(* IEC 61131-3 sources: deprecated-refusr-repo/samples (part 25) *)

(* ---- RND-EXPR_calms-hitch-chips.st ---- *)
(*
This code implements a randomly grown symbolic expression:

((((!(xor(xor(IN37 & (IN27 | ((IN12 & IN24) | (xor(xor(IN9, IN8), IN8)))), (((IN7 & IN10) | (IN4 | IN33)) & IN19) & (xor(xor(!(xor(xor(IN45, IN17), IN10)), !(IN49)), (IN17 & IN40) & (IN49 & IN27)))), (IN29 & (!(xor(xor(IN44, IN27), IN49)))) & IN44))) & (xor(xor((xor(xor(IN25 & ((IN10 | IN28) & IN1), xor(xor(!(!(IN7)), IN13 | (IN39 & IN48)), !(IN32 | IN22))), IN12 & IN3)) & (((!(IN1 & true)) | (IN40 & (!(IN33)))) & ((!(!(IN39))) & ((IN31 | IN24) & IN12))), ((!(IN45)) | ((IN39 | (IN21 | IN31)) | IN2)) | (xor(xor(xor(xor(!(IN20 & IN8), xor(xor(xor(xor(IN3, IN22), IN23), !(IN26)), IN36 & IN23)), !(IN7 | IN30)), (IN12 & (IN40 & IN39)) & (!(IN11 | IN36))), IN48 | IN27))), (!((!(false | IN8)) & ((IN41 & IN46) | (!(IN10))))) & ((!((xor(xor(IN49, IN16), IN2)) | (xor(xor(IN1, IN43), IN14)))) & (!(xor(xor(true & IN26, !(IN43)), xor(xor(IN50, IN38), IN31)))))))) | (((xor(xor(IN15 & (((!(IN16)) & (xor(xor(IN17, IN4), IN20))) & (!(IN23))), (!(xor(xor(false & IN33, xor(xor(IN43, IN26), IN5)), IN34 | IN13))) | (!((xor(xor(IN34, IN42), IN26)) | (!(IN14))))), (((IN10 | IN35) & (IN3 & IN6)) | ((!(IN24)) & (xor(xor(IN26, IN21), IN4)))) | (!(!(IN39 & IN43))))) & (IN6 | ((!(!(xor(xor(IN12, IN16), IN44)))) & IN38))) | (xor(xor(IN25, (xor(xor(xor(xor(!(IN8 & IN48), xor(xor(IN32 | IN43, IN16 | IN16), IN36 | IN46)), xor(xor(IN47, !(IN48)), IN35 | IN43)), xor(xor((IN45 | true) | (!(IN18)), IN13 | (xor(xor(IN5, IN40), IN37))), (!(IN32)) | (!(IN30)))), ((IN6 & IN50) | (IN12 | IN40)) | (xor(xor(!(IN26), xor(xor(IN28, IN10), IN19)), IN30 | IN9)))) & (!(((IN36 & IN40) & (!(IN27))) & (xor(xor(IN36 & true, IN6 | IN2), xor(xor(IN17, IN35), IN35)))))), xor(xor((!(!(IN3 | IN2))) & (!(!(IN13))), IN28), ((!(IN49 & IN49)) | (!(IN7 & IN22))) & (!((IN34 & IN14) & (IN33 | IN12)))))))) & (!(IN3))) & ((!((xor(xor(IN17, !((((IN49 & IN26) | (xor(xor(IN36, IN25), false))) & (xor(xor(IN5 & false, !(IN35)), !(IN50)))) & (!(!(IN6 | IN36))))), !(IN48 & IN8))) & ((xor(xor((!((xor(xor(IN33, IN8), IN42)) | (!(IN38)))) & (xor(xor(!(!(IN31)), xor(xor(IN29, !(IN19)), IN30 & IN32)), xor(xor(IN21, IN19), IN26 | IN33))), (xor(xor((!(IN43)) | (IN50 | IN48), !(!(IN4))), (IN46 | IN17) | (IN30 & IN5))) | ((xor(xor(!(IN13), !(IN13)), xor(xor(IN47, IN28), IN11))) & (xor(xor(!(IN34), IN1 & IN9), IN18 | IN18)))), !(!(!(xor(xor(IN27, IN9), IN50)))))) | (xor(xor(xor(xor(((IN38 | IN16) & (xor(xor(IN41, IN33), IN19))) | (!(xor(xor(IN24, IN1), IN26))), IN22 | ((!(IN32)) | (IN39 & IN2))), ((xor(xor(IN29, IN31), IN5)) & (IN28 | IN27)) & IN20), IN48 & (!((!(IN49)) | (IN30 & IN43)))), IN17 | (((xor(xor(IN21, IN47), IN26)) & (IN28 | false)) | (!(IN31 & false)))))))) & (xor(xor((xor(xor(!((!(!(IN14 & IN46))) & IN35), IN1 | (((!(!(IN20))) & (xor(xor(IN14 & IN29, IN28 & IN20), IN24 & IN18))) & (!(!(IN15 & IN16))))), (xor(xor(((xor(xor(IN14, IN48), IN24)) & (xor(xor(IN5, IN43), IN5))) | ((IN22 | IN46) | (IN44 & IN8)), !((xor(xor(IN50, IN32), IN48)) | (xor(xor(IN28, IN47), IN47)))), (!(xor(xor(IN20, IN39), IN43))) | (!(IN21 & IN17)))) & ((((IN36 | IN24) & (IN9 & IN28)) & IN6) & (true & IN18)))) & ((xor(xor((xor(xor(!(xor(xor(IN44, IN27), IN50)), IN14), IN44)) | (!(!(xor(xor(IN15, IN29), IN24)))), (IN7 & (IN34 | (xor(xor(IN14, IN19), IN41)))) | (((IN10 & IN43) | (IN32 | IN38)) & ((IN5 & IN35) | IN1))), IN43)) | (xor(xor(IN45, xor(xor(true | (!(IN49 | IN18)), IN33 & (!(IN5 & IN13))), IN43)), IN5))), (!((IN23 | ((!(IN45 | IN31)) & IN9)) | (xor(xor(!((IN27 | IN21) & (!(IN26))), !(IN27)), ((IN48 & IN48) & (xor(xor(IN37, IN41), IN13))) & IN49)))) | (((!(((!(IN15)) | (xor(xor(IN1, IN25), IN6))) | IN46)) | IN13) & ((IN18 | (xor(xor(IN14 & (!(IN35)), xor(xor(xor(xor(IN40, IN41), IN23), xor(xor(IN6, IN18), IN22)), IN10)), IN35))) | (!(((IN34 & IN11) & (IN46 & IN43)) & (xor(xor(IN31, IN25 | IN32), xor(xor(IN35, IN11), IN9)))))))), !(((xor(xor(xor(xor(IN39, IN42 | (xor(xor(IN33, IN4), IN29))), IN24 & (!(IN45))), (xor(xor(!(IN11), IN39 & false), IN35)) & ((xor(xor(IN12, IN35), IN44)) & IN30)), xor(xor(IN23, !(!(IN25))), !(IN25 & IN14)))) & (IN24 | ((xor(xor(IN4, !(IN27)), IN28 | IN44)) | (xor(xor(IN44 & IN22, IN44 | IN50), IN44))))) | (!((xor(xor(!(IN23), (xor(xor(IN24, IN35), IN27)) & (IN27 | IN14)), (!(IN37)) & (!(IN27)))) & ((xor(xor(IN24 & IN33, IN3), !(IN16))) & ((IN12 | IN39) & IN25))))))))

*)

FUNCTION_BLOCK F_CollectInput
  VAR_IN_OUT
      Data : ARRAY[1..50] OF BOOL;
  END_VAR
  VAR_INPUT
      TICK  : BOOL := 0;
      IN1   : BOOL := 0;
      IN2   : BOOL := 0;
      IN3   : BOOL := 0;
      IN4   : BOOL := 0;
      IN5   : BOOL := 0;
      RESET : BOOL := FALSE;
  END_VAR
  VAR_OUTPUT
      Finished : BOOL;
  END_VAR
  VAR
      j    : USINT := 1;
      tock : BOOL  := 0;
  END_VAR
  IF NOT RESET AND tock = NOT TICK THEN
      Data[j]   := IN1;
      Data[j+1] := IN2;
      Data[j+2] := IN3;
      Data[j+3] := IN4;
      Data[j+4] := IN5;
      j := j + 5;
      tock := TICK;
  ELSE
      j := 1;
      tock := 0;
  END_IF;
  Finished := (j > 50);
END_FUNCTION_BLOCK

PROGRAM Boiler
  VAR
    Data  : ARRAY[1..50] OF BOOL;
    Ready : BOOL;
    CollectInput : F_CollectInput;
  END_VAR
  VAR
    TICK     AT %IX1.0 : BOOL;
    IN1      AT %IX0.3 : BOOL;
    IN2      AT %IX0.4 : BOOL;
    IN3      AT %IX0.5 : BOOL;
    IN4      AT %IX0.6 : BOOL;
    IN5      AT %IX0.7 : BOOL;
    OutReady AT %QX0.0 : BOOL := FALSE;
    FeedNext AT %QX0.1 : BOOL := FALSE;
    Out      AT %QX0.2 : BOOL;
  END_VAR
  CollectInput(TICK:=TICK, IN1:=IN1, IN2:=IN2, IN3:=IN3, IN4:=IN4, IN5:=IN5);
  Ready := CollectInput.Finished;
  FeedNext := 1;
  IF Ready THEN
    Out := (((((NOT (((Data[37] AND (Data[27] OR ((Data[12] AND Data[24]) OR ((Data[9] XOR Data[8]) XOR Data[8])))) XOR ((((Data[7] AND Data[10]) OR (Data[4] OR Data[33])) AND Data[19]) AND (((NOT ((Data[45] XOR Data[17]) XOR Data[10])) XOR (NOT Data[49])) XOR ((Data[17] AND Data[40]) AND (Data[49] AND Data[27]))))) XOR ((Data[29] AND (NOT ((Data[44] XOR Data[27]) XOR Data[49]))) AND Data[44]))) AND ((((((Data[25] AND ((Data[10] OR Data[28]) AND Data[1])) XOR (((NOT (NOT Data[7])) XOR (Data[13] OR (Data[39] AND Data[48]))) XOR (NOT (Data[32] OR Data[22])))) XOR (Data[12] AND Data[3])) AND (((NOT (Data[1] AND TRUE)) OR (Data[40] AND (NOT Data[33]))) AND ((NOT (NOT Data[39])) AND ((Data[31] OR Data[24]) AND Data[12])))) XOR (((NOT Data[45]) OR ((Data[39] OR (Data[21] OR Data[31])) OR Data[2])) OR (((((NOT (Data[20] AND Data[8])) XOR ((((Data[3] XOR Data[22]) XOR Data[23]) XOR (NOT Data[26])) XOR (Data[36] AND Data[23]))) XOR (NOT (Data[7] OR Data[30]))) XOR ((Data[12] AND (Data[40] AND Data[39])) AND (NOT (Data[11] OR Data[36])))) XOR (Data[48] OR Data[27])))) XOR ((NOT ((NOT (FALSE OR Data[8])) AND ((Data[41] AND Data[46]) OR (NOT Data[10])))) AND ((NOT (((Data[49] XOR Data[16]) XOR Data[2]) OR ((Data[1] XOR Data[43]) XOR Data[14]))) AND (NOT (((TRUE AND Data[26]) XOR (NOT Data[43])) XOR ((Data[50] XOR Data[38]) XOR Data[31]))))))) OR (((((Data[15] AND (((NOT Data[16]) AND ((Data[17] XOR Data[4]) XOR Data[20])) AND (NOT Data[23]))) XOR ((NOT (((FALSE AND Data[33]) XOR ((Data[43] XOR Data[26]) XOR Data[5])) XOR (Data[34] OR Data[13]))) OR (NOT (((Data[34] XOR Data[42]) XOR Data[26]) OR (NOT Data[14]))))) XOR ((((Data[10] OR Data[35]) AND (Data[3] AND Data[6])) OR ((NOT Data[24]) AND ((Data[26] XOR Data[21]) XOR Data[4]))) OR (NOT (NOT (Data[39] AND Data[43]))))) AND (Data[6] OR ((NOT (NOT ((Data[12] XOR Data[16]) XOR Data[44]))) AND Data[38]))) OR ((Data[25] XOR ((((((NOT (Data[8] AND Data[48])) XOR (((Data[32] OR Data[43]) XOR (Data[16] OR Data[16])) XOR (Data[36] OR Data[46]))) XOR ((Data[47] XOR (NOT Data[48])) XOR (Data[35] OR Data[43]))) XOR ((((Data[45] OR TRUE) OR (NOT Data[18])) XOR (Data[13] OR ((Data[5] XOR Data[40]) XOR Data[37]))) XOR ((NOT Data[32]) OR (NOT Data[30])))) XOR (((Data[6] AND Data[50]) OR (Data[12] OR Data[40])) OR (((NOT Data[26]) XOR ((Data[28] XOR Data[10]) XOR Data[19])) XOR (Data[30] OR Data[9])))) AND (NOT (((Data[36] AND Data[40]) AND (NOT Data[27])) AND (((Data[36] AND TRUE) XOR (Data[6] OR Data[2])) XOR ((Data[17] XOR Data[35]) XOR Data[35])))))) XOR ((((NOT (NOT (Data[3] OR Data[2]))) AND (NOT (NOT Data[13]))) XOR Data[28]) XOR (((NOT (Data[49] AND Data[49])) OR (NOT (Data[7] AND Data[22]))) AND (NOT ((Data[34] AND Data[14]) AND (Data[33] OR Data[12])))))))) AND (NOT Data[3])) AND ((NOT (((Data[17] XOR (NOT ((((Data[49] AND Data[26]) OR ((Data[36] XOR Data[25]) XOR FALSE)) AND (((Data[5] AND FALSE) XOR (NOT Data[35])) XOR (NOT Data[50]))) AND (NOT (NOT (Data[6] OR Data[36])))))) XOR (NOT (Data[48] AND Data[8]))) AND (((((NOT (((Data[33] XOR Data[8]) XOR Data[42]) OR (NOT Data[38]))) AND (((NOT (NOT Data[31])) XOR ((Data[29] XOR (NOT Data[19])) XOR (Data[30] AND Data[32]))) XOR ((Data[21] XOR Data[19]) XOR (Data[26] OR Data[33])))) XOR (((((NOT Data[43]) OR (Data[50] OR Data[48])) XOR (NOT (NOT Data[4]))) XOR ((Data[46] OR Data[17]) OR (Data[30] AND Data[5]))) OR ((((NOT Data[13]) XOR (NOT Data[13])) XOR ((Data[47] XOR Data[28]) XOR Data[11])) AND (((NOT Data[34]) XOR (Data[1] AND Data[9])) XOR (Data[18] OR Data[18]))))) XOR (NOT (NOT (NOT ((Data[27] XOR Data[9]) XOR Data[50]))))) OR (((((((Data[38] OR Data[16]) AND ((Data[41] XOR Data[33]) XOR Data[19])) OR (NOT ((Data[24] XOR Data[1]) XOR Data[26]))) XOR (Data[22] OR ((NOT Data[32]) OR (Data[39] AND Data[2])))) XOR ((((Data[29] XOR Data[31]) XOR Data[5]) AND (Data[28] OR Data[27])) AND Data[20])) XOR (Data[48] AND (NOT ((NOT Data[49]) OR (Data[30] AND Data[43]))))) XOR (Data[17] OR ((((Data[21] XOR Data[47]) XOR Data[26]) AND (Data[28] OR FALSE)) OR (NOT (Data[31] AND FALSE)))))))) AND ((((((NOT ((NOT (NOT (Data[14] AND Data[46]))) AND Data[35])) XOR (Data[1] OR (((NOT (NOT Data[20])) AND (((Data[14] AND Data[29]) XOR (Data[28] AND Data[20])) XOR (Data[24] AND Data[18]))) AND (NOT (NOT (Data[15] AND Data[16])))))) XOR (((((((Data[14] XOR Data[48]) XOR Data[24]) AND ((Data[5] XOR Data[43]) XOR Data[5])) OR ((Data[22] OR Data[46]) OR (Data[44] AND Data[8]))) XOR (NOT (((Data[50] XOR Data[32]) XOR Data[48]) OR ((Data[28] XOR Data[47]) XOR Data[47])))) XOR ((NOT ((Data[20] XOR Data[39]) XOR Data[43])) OR (NOT (Data[21] AND Data[17])))) AND ((((Data[36] OR Data[24]) AND (Data[9] AND Data[28])) AND Data[6]) AND (TRUE AND Data[18])))) AND (((((((NOT ((Data[44] XOR Data[27]) XOR Data[50])) XOR Data[14]) XOR Data[44]) OR (NOT (NOT ((Data[15] XOR Data[29]) XOR Data[24])))) XOR ((Data[7] AND (Data[34] OR ((Data[14] XOR Data[19]) XOR Data[41]))) OR (((Data[10] AND Data[43]) OR (Data[32] OR Data[38])) AND ((Data[5] AND Data[35]) OR Data[1])))) XOR Data[43]) OR ((Data[45] XOR (((TRUE OR (NOT (Data[49] OR Data[18]))) XOR (Data[33] AND (NOT (Data[5] AND Data[13])))) XOR Data[43])) XOR Data[5]))) XOR ((NOT ((Data[23] OR ((NOT (Data[45] OR Data[31])) AND Data[9])) OR (((NOT ((Data[27] OR Data[21]) AND (NOT Data[26]))) XOR (NOT Data[27])) XOR (((Data[48] AND Data[48]) AND ((Data[37] XOR Data[41]) XOR Data[13])) AND Data[49])))) OR (((NOT (((NOT Data[15]) OR ((Data[1] XOR Data[25]) XOR Data[6])) OR Data[46])) OR Data[13]) AND ((Data[18] OR (((Data[14] AND (NOT Data[35])) XOR ((((Data[40] XOR Data[41]) XOR Data[23]) XOR ((Data[6] XOR Data[18]) XOR Data[22])) XOR Data[10])) XOR Data[35])) OR (NOT (((Data[34] AND Data[11]) AND (Data[46] AND Data[43])) AND ((Data[31] XOR (Data[25] OR Data[32])) XOR ((Data[35] XOR Data[11]) XOR Data[9])))))))) XOR (NOT ((((((Data[39] XOR (Data[42] OR ((Data[33] XOR Data[4]) XOR Data[29]))) XOR (Data[24] AND (NOT Data[45]))) XOR ((((NOT Data[11]) XOR (Data[39] AND FALSE)) XOR Data[35]) AND (((Data[12] XOR Data[35]) XOR Data[44]) AND Data[30]))) XOR ((Data[23] XOR (NOT (NOT Data[25]))) XOR (NOT (Data[25] AND Data[14])))) AND (Data[24] OR (((Data[4] XOR (NOT Data[27])) XOR (Data[28] OR Data[44])) OR (((Data[44] AND Data[22]) XOR (Data[44] OR Data[50])) XOR Data[44])))) OR (NOT ((((NOT Data[23]) XOR (((Data[24] XOR Data[35]) XOR Data[27]) AND (Data[27] OR Data[14]))) XOR ((NOT Data[37]) AND (NOT Data[27]))) AND ((((Data[24] AND Data[33]) XOR Data[3]) XOR (NOT Data[16])) AND ((Data[12] OR Data[39]) AND Data[25])))))))));
    OutReady := 1;
    CollectInput(RESET:=TRUE);
  END_IF;
END_PROGRAM

CONFIGURATION Config0
  RESOURCE Res0 ON PLC
    TASK task0(INTERVAL := T#20ms,PRIORITY := 0);
    PROGRAM instance0 WITH task0 : Boiler;
  END_RESOURCE
END_CONFIGURATION

(* ---- RND-EXPR_celeb-candy-degas.st ---- *)
(*
This code implements a randomly grown symbolic expression:

!(xor(xor(!(!(((IN43 & ((xor(xor(IN28 | IN19, !(IN27)), IN33 | IN34)) & (xor(xor(xor(xor(IN27, IN17), IN17), xor(xor(true, IN6), IN43)), xor(xor(IN12, IN24), IN27))))) | IN22) & ((!(xor(xor(IN48, true), IN11))) | (((!(IN32)) | (!(IN3 | IN3))) | ((!(IN10)) | ((IN29 | IN6) | IN19)))))), xor(xor(xor(xor(IN26, !(IN24)), ((IN50 | ((xor(xor(IN4 & IN32, xor(xor(IN29, IN44), IN1)), IN25 & IN41)) | ((IN17 | IN36) & (xor(xor(IN10, IN2), IN16))))) & ((!(!(IN10))) | (!((!(IN48)) | (IN8 | IN19))))) | (!(!(((IN1 | IN6) | IN48) | (IN15 & IN7))))), ((xor(xor(xor(xor((xor(xor(!(IN39), !(IN1)), IN33 | IN10)) | IN5, xor(xor((IN21 | IN15) & (xor(xor(IN35, IN25), IN41)), (IN18 | IN2) & IN21), (IN2 | IN3) & (!(IN39)))), xor(xor((IN36 | IN33) | (!(IN14)), !(!(IN39))), !(IN16 & IN8))), IN15), (xor(xor(xor(xor(IN6 | IN24, xor(xor(IN49, IN14), IN21)), xor(xor(IN13, IN16), IN43)), !(xor(xor(IN23, IN10), IN19))), xor(xor(IN6 | IN31, xor(xor(IN40, IN38), IN29)), IN43))) & ((IN38 | (!(IN28))) | ((xor(xor(IN33, IN34), IN36)) & IN13)))) | IN42) | (((xor(xor((xor(xor(IN4, xor(xor(IN6, IN6), IN31)), !(IN21))) | (!(xor(xor(IN21, false), IN15))), IN17), ((xor(xor(false, IN5), IN47)) & (xor(xor(IN49, IN19), IN41))) & (xor(xor(!(IN38), IN8 | IN34), IN15 & IN16)))) | IN18) & ((IN38 & (IN28 & IN1)) | (xor(xor((IN10 | (!(IN33))) | IN45, (!(IN6 & IN5)) & ((!(IN3)) | IN19)), xor(xor(xor(xor(!(IN28), IN16 | IN32), IN2 | IN9), (IN39 | IN36) & (!(IN41))), (!(IN26)) | (!(IN47)))))))), xor(xor(!(((((IN14 | false) & IN34) & (IN23 & (IN13 | IN3))) & (((IN45 & IN1) | (xor(xor(IN22, IN35), IN4))) | (IN2 & IN25))) | IN26), xor(xor(xor(xor((IN2 & (xor(xor(xor(xor(IN4, IN28), IN34), IN3 & IN28), IN24 | IN22))) | IN16, (xor(xor(!(IN26 & IN50), !(IN13 | IN37)), !(IN35))) | (((!(IN35)) & IN24) & (!(IN24 & IN12)))), xor(xor(!((!(IN10)) | (IN9 | IN28)), ((IN35 | IN46) & IN4) | (xor(xor(false, xor(xor(IN22, IN24), IN1)), IN22 | IN21))), ((IN29 & IN33) | (xor(xor(false, IN45), IN26))) | IN30)), !(IN19)), xor(xor(false, !((xor(xor(IN22 | IN45, xor(xor(IN12, true), IN19)), IN35 & IN24)) | (!(IN46)))), IN50))), IN39))), xor(xor(IN12 & (xor(xor(!(xor(xor(((xor(xor(IN31, IN35), IN20)) & (!(IN37))) & ((xor(xor(IN15, IN38), IN12)) & (xor(xor(IN19, IN42), IN31))), ((IN9 & IN29) | (!(IN16))) & IN5), ((xor(xor(IN21, IN25), IN21)) | (IN21 | IN17)) & (!(!(IN42))))), xor(xor((xor(xor(IN12, !(xor(xor(IN48, true), IN39))), (IN21 | IN43) | (IN12 | true))) | ((xor(xor(IN31 | IN44, IN18 & IN48), xor(xor(IN11, IN35), IN21))) & (xor(xor(xor(xor(IN25, IN40), IN10), IN13 & true), xor(xor(IN47, IN22), IN21)))), (xor(xor((!(IN36)) & (IN29 & IN15), IN35), IN46)) & (!(IN32))), !(!((!(IN27)) & (!(IN36)))))), (!(((IN1 & IN21) | (!(IN45))) | ((IN23 & IN32) | IN41))) & (xor(xor(xor(xor(IN40, (!(IN32)) & (IN20 | IN20)), xor(xor(xor(xor(IN26, IN20), IN50), IN8 & IN49), IN4 & IN21)), ((xor(xor(IN25, IN6), IN39)) & (IN10 & IN16)) & (xor(xor(IN14 & IN33, IN3 & IN21), IN28 | IN18))), IN13)))), xor(xor(xor(xor(!((!(xor(xor(IN29 & IN49, IN32), xor(xor(IN15, IN21), IN3)))) | (!(IN49 & (xor(xor(IN23, IN40), IN49))))), (xor(xor(((!(IN49)) & (IN28 & IN26)) & IN23, ((IN43 & IN42) | IN39) & (!(IN38 | IN22))), (!(IN17)) & IN50)) & ((xor(xor(xor(xor(xor(xor(IN50, IN5), IN38), xor(xor(IN49, IN32), IN31)), !(IN18)), IN11), (!(IN6)) | IN38)) & IN48)), IN50 & IN22), ((xor(xor(IN31 & true, (!(IN47 & IN18)) | (!(!(IN48)))), (!(!(IN50))) | IN28)) | ((!((IN7 | IN24) | (IN4 | IN44))) | (xor(xor(!(IN9), IN39), (false & IN12) | (IN26 & IN50))))) & IN35), !((!(xor(xor(IN7, (!(IN38)) & (IN38 | IN17)), xor(xor(xor(xor(IN49, IN21), IN35), IN17 & IN21), xor(xor(IN45, IN26), IN29))))) | ((IN36 & (xor(xor(xor(xor(IN11, IN31), IN32), IN46 & IN49), !(IN2)))) & (!(!(IN24))))))), xor(xor(xor(xor(!(IN1 & IN12), (!(xor(xor(xor(xor(!(IN44), IN35), IN41 | IN16), xor(xor(IN39 & IN2, !(IN19)), IN25)), !(IN21)))) | ((((xor(xor(IN27, IN33), false)) & IN29) | ((IN4 & IN18) | (IN2 | IN36))) & IN46)), (IN23 | (!(IN13))) & (!((true & (IN42 & IN20)) | (xor(xor(!(IN12), IN7 | true), IN1 | IN14))))), IN21), !(!(IN29))))))

*)

FUNCTION_BLOCK F_CollectInput
  VAR_IN_OUT
      Data : ARRAY[1..50] OF BOOL;
  END_VAR
  VAR_INPUT
      TICK  : BOOL := 0;
      IN1   : BOOL := 0;
      IN2   : BOOL := 0;
      IN3   : BOOL := 0;
      IN4   : BOOL := 0;
      IN5   : BOOL := 0;
      RESET : BOOL := FALSE;
  END_VAR
  VAR_OUTPUT
      Finished : BOOL;
  END_VAR
  VAR
      j    : USINT := 1;
      tock : BOOL  := 0;
  END_VAR
  IF NOT RESET AND tock = NOT TICK THEN
      Data[j]   := IN1;
      Data[j+1] := IN2;
      Data[j+2] := IN3;
      Data[j+3] := IN4;
      Data[j+4] := IN5;
      j := j + 5;
      tock := TICK;
  ELSE
      j := 1;
      tock := 0;
  END_IF;
  Finished := (j > 50);
END_FUNCTION_BLOCK

PROGRAM Boiler
  VAR
    Data  : ARRAY[1..50] OF BOOL;
    Ready : BOOL;
    CollectInput : F_CollectInput;
  END_VAR
  VAR
    TICK     AT %IX1.0 : BOOL;
    IN1      AT %IX0.3 : BOOL;
    IN2      AT %IX0.4 : BOOL;
    IN3      AT %IX0.5 : BOOL;
    IN4      AT %IX0.6 : BOOL;
    IN5      AT %IX0.7 : BOOL;
    OutReady AT %QX0.0 : BOOL := FALSE;
    FeedNext AT %QX0.1 : BOOL := FALSE;
    Out      AT %QX0.2 : BOOL;
  END_VAR
  CollectInput(TICK:=TICK, IN1:=IN1, IN2:=IN2, IN3:=IN3, IN4:=IN4, IN5:=IN5);
  Ready := CollectInput.Finished;
  FeedNext := 1;
  IF Ready THEN
    Out := (NOT (((NOT (NOT (((Data[43] AND ((((Data[28] OR Data[19]) XOR (NOT Data[27])) XOR (Data[33] OR Data[34])) AND ((((Data[27] XOR Data[17]) XOR Data[17]) XOR ((TRUE XOR Data[6]) XOR Data[43])) XOR ((Data[12] XOR Data[24]) XOR Data[27])))) OR Data[22]) AND ((NOT ((Data[48] XOR TRUE) XOR Data[11])) OR (((NOT Data[32]) OR (NOT (Data[3] OR Data[3]))) OR ((NOT Data[10]) OR ((Data[29] OR Data[6]) OR Data[19]))))))) XOR ((((Data[26] XOR (NOT Data[24])) XOR (((Data[50] OR ((((Data[4] AND Data[32]) XOR ((Data[29] XOR Data[44]) XOR Data[1])) XOR (Data[25] AND Data[41])) OR ((Data[17] OR Data[36]) AND ((Data[10] XOR Data[2]) XOR Data[16])))) AND ((NOT (NOT Data[10])) OR (NOT ((NOT Data[48]) OR (Data[8] OR Data[19]))))) OR (NOT (NOT (((Data[1] OR Data[6]) OR Data[48]) OR (Data[15] AND Data[7])))))) XOR ((((((((((NOT Data[39]) XOR (NOT Data[1])) XOR (Data[33] OR Data[10])) OR Data[5]) XOR ((((Data[21] OR Data[15]) AND ((Data[35] XOR Data[25]) XOR Data[41])) XOR ((Data[18] OR Data[2]) AND Data[21])) XOR ((Data[2] OR Data[3]) AND (NOT Data[39])))) XOR ((((Data[36] OR Data[33]) OR (NOT Data[14])) XOR (NOT (NOT Data[39]))) XOR (NOT (Data[16] AND Data[8])))) XOR Data[15]) XOR ((((((Data[6] OR Data[24]) XOR ((Data[49] XOR Data[14]) XOR Data[21])) XOR ((Data[13] XOR Data[16]) XOR Data[43])) XOR (NOT ((Data[23] XOR Data[10]) XOR Data[19]))) XOR (((Data[6] OR Data[31]) XOR ((Data[40] XOR Data[38]) XOR Data[29])) XOR Data[43])) AND ((Data[38] OR (NOT Data[28])) OR (((Data[33] XOR Data[34]) XOR Data[36]) AND Data[13])))) OR Data[42]) OR (((((((Data[4] XOR ((Data[6] XOR Data[6]) XOR Data[31])) XOR (NOT Data[21])) OR (NOT ((Data[21] XOR FALSE) XOR Data[15]))) XOR Data[17]) XOR ((((FALSE XOR Data[5]) XOR Data[47]) AND ((Data[49] XOR Data[19]) XOR Data[41])) AND (((NOT Data[38]) XOR (Data[8] OR Data[34])) XOR (Data[15] AND Data[16])))) OR Data[18]) AND ((Data[38] AND (Data[28] AND Data[1])) OR ((((Data[10] OR (NOT Data[33])) OR Data[45]) XOR ((NOT (Data[6] AND Data[5])) AND ((NOT Data[3]) OR Data[19]))) XOR (((((NOT Data[28]) XOR (Data[16] OR Data[32])) XOR (Data[2] OR Data[9])) XOR ((Data[39] OR Data[36]) AND (NOT Data[41]))) XOR ((NOT Data[26]) OR (NOT Data[47])))))))) XOR (((NOT (((((Data[14] OR FALSE) AND Data[34]) AND (Data[23] AND (Data[13] OR Data[3]))) AND (((Data[45] AND Data[1]) OR ((Data[22] XOR Data[35]) XOR Data[4])) OR (Data[2] AND Data[25]))) OR Data[26])) XOR ((((((Data[2] AND ((((Data[4] XOR Data[28]) XOR Data[34]) XOR (Data[3] AND Data[28])) XOR (Data[24] OR Data[22]))) OR Data[16]) XOR ((((NOT (Data[26] AND Data[50])) XOR (NOT (Data[13] OR Data[37]))) XOR (NOT Data[35])) OR (((NOT Data[35]) AND Data[24]) AND (NOT (Data[24] AND Data[12]))))) XOR (((NOT ((NOT Data[10]) OR (Data[9] OR Data[28]))) XOR (((Data[35] OR Data[46]) AND Data[4]) OR ((FALSE XOR ((Data[22] XOR Data[24]) XOR Data[1])) XOR (Data[22] OR Data[21])))) XOR (((Data[29] AND Data[33]) OR ((FALSE XOR Data[45]) XOR Data[26])) OR Data[30]))) XOR (NOT Data[19])) XOR ((FALSE XOR (NOT ((((Data[22] OR Data[45]) XOR ((Data[12] XOR TRUE) XOR Data[19])) XOR (Data[35] AND Data[24])) OR (NOT Data[46])))) XOR Data[50]))) XOR Data[39]))) XOR (((Data[12] AND (((NOT ((((((Data[31] XOR Data[35]) XOR Data[20]) AND (NOT Data[37])) AND (((Data[15] XOR Data[38]) XOR Data[12]) AND ((Data[19] XOR Data[42]) XOR Data[31]))) XOR (((Data[9] AND Data[29]) OR (NOT Data[16])) AND Data[5])) XOR ((((Data[21] XOR Data[25]) XOR Data[21]) OR (Data[21] OR Data[17])) AND (NOT (NOT Data[42]))))) XOR (((((Data[12] XOR (NOT ((Data[48] XOR TRUE) XOR Data[39]))) XOR ((Data[21] OR Data[43]) OR (Data[12] OR TRUE))) OR ((((Data[31] OR Data[44]) XOR (Data[18] AND Data[48])) XOR ((Data[11] XOR Data[35]) XOR Data[21])) AND ((((Data[25] XOR Data[40]) XOR Data[10]) XOR (Data[13] AND TRUE)) XOR ((Data[47] XOR Data[22]) XOR Data[21])))) XOR (((((NOT Data[36]) AND (Data[29] AND Data[15])) XOR Data[35]) XOR Data[46]) AND (NOT Data[32]))) XOR (NOT (NOT ((NOT Data[27]) AND (NOT Data[36])))))) XOR ((NOT (((Data[1] AND Data[21]) OR (NOT Data[45])) OR ((Data[23] AND Data[32]) OR Data[41]))) AND ((((Data[40] XOR ((NOT Data[32]) AND (Data[20] OR Data[20]))) XOR ((((Data[26] XOR Data[20]) XOR Data[50]) XOR (Data[8] AND Data[49])) XOR (Data[4] AND Data[21]))) XOR ((((Data[25] XOR Data[6]) XOR Data[39]) AND (Data[10] AND Data[16])) AND (((Data[14] AND Data[33]) XOR (Data[3] AND Data[21])) XOR (Data[28] OR Data[18])))) XOR Data[13])))) XOR (((((NOT ((NOT (((Data[29] AND Data[49]) XOR Data[32]) XOR ((Data[15] XOR Data[21]) XOR Data[3]))) OR (NOT (Data[49] AND ((Data[23] XOR Data[40]) XOR Data[49]))))) XOR ((((((NOT Data[49]) AND (Data[28] AND Data[26])) AND Data[23]) XOR (((Data[43] AND Data[42]) OR Data[39]) AND (NOT (Data[38] OR Data[22])))) XOR ((NOT Data[17]) AND Data[50])) AND (((((((Data[50] XOR Data[5]) XOR Data[38]) XOR ((Data[49] XOR Data[32]) XOR Data[31])) XOR (NOT Data[18])) XOR Data[11]) XOR ((NOT Data[6]) OR Data[38])) AND Data[48]))) XOR (Data[50] AND Data[22])) XOR (((((Data[31] AND TRUE) XOR ((NOT (Data[47] AND Data[18])) OR (NOT (NOT Data[48])))) XOR ((NOT (NOT Data[50])) OR Data[28])) OR ((NOT ((Data[7] OR Data[24]) OR (Data[4] OR Data[44]))) OR (((NOT Data[9]) XOR Data[39]) XOR ((FALSE AND Data[12]) OR (Data[26] AND Data[50]))))) AND Data[35])) XOR (NOT ((NOT ((Data[7] XOR ((NOT Data[38]) AND (Data[38] OR Data[17]))) XOR ((((Data[49] XOR Data[21]) XOR Data[35]) XOR (Data[17] AND Data[21])) XOR ((Data[45] XOR Data[26]) XOR Data[29])))) OR ((Data[36] AND ((((Data[11] XOR Data[31]) XOR Data[32]) XOR (Data[46] AND Data[49])) XOR (NOT Data[2]))) AND (NOT (NOT Data[24]))))))) XOR (((((NOT (Data[1] AND Data[12])) XOR ((NOT (((((NOT Data[44]) XOR Data[35]) XOR (Data[41] OR Data[16])) XOR (((Data[39] AND Data[2]) XOR (NOT Data[19])) XOR Data[25])) XOR (NOT Data[21]))) OR (((((Data[27] XOR Data[33]) XOR FALSE) AND Data[29]) OR ((Data[4] AND Data[18]) OR (Data[2] OR Data[36]))) AND Data[46]))) XOR ((Data[23] OR (NOT Data[13])) AND (NOT ((TRUE AND (Data[42] AND Data[20])) OR (((NOT Data[12]) XOR (Data[7] OR TRUE)) XOR (Data[1] OR Data[14])))))) XOR Data[21]) XOR (NOT (NOT Data[29]))))));
    OutReady := 1;
    CollectInput(RESET:=TRUE);
  END_IF;
END_PROGRAM

CONFIGURATION Config0
  RESOURCE Res0 ON PLC
    TASK task0(INTERVAL := T#20ms,PRIORITY := 0);
    PROGRAM instance0 WITH task0 : Boiler;
  END_RESOURCE
END_CONFIGURATION

(* ---- RND-EXPR_endue-lawns-artsy.st ---- *)
(*
This code implements a randomly grown symbolic expression:

xor(xor(xor(xor(!(xor(xor(IN45, xor(xor((((xor(xor(IN19 & IN49, IN3 & IN10), !(IN13))) | IN18) & (IN2 | ((xor(xor(IN32, IN39), IN18)) | IN26))) | (!(((IN23 & IN4) & (!(IN25))) & (xor(xor(!(IN15), xor(xor(IN16, IN30), IN44)), xor(xor(IN26, true), IN50))))), !(((!(xor(xor(IN16, IN38), IN11))) | (IN17 | (!(IN22)))) | (!(!(!(IN31)))))), (((!(IN2)) & (!(IN49 | IN20))) & (xor(xor(IN27 & (xor(xor(IN47, IN2), true)), (IN21 | IN9) | IN35), IN15 | (!(IN16))))) & ((!(!(!(IN17)))) | (!(xor(xor(IN48, IN15 & IN19), xor(xor(IN13, IN36), IN25))))))), xor(xor(IN14 & (xor(xor(xor(xor((IN38 & IN38) & (IN45 | IN6), (IN12 & IN4) | (IN47 | IN26)), xor(xor(xor(xor(IN2, IN1), IN42), IN41 | IN2), IN43 | IN10)), (!(IN24 | IN39)) & (xor(xor(IN35 | IN36, xor(xor(IN4, IN46), IN47)), IN50))), (!(xor(xor(IN28, IN30), IN39))) & ((xor(xor(IN49, false), IN31)) & (IN28 | IN47)))), IN15), !(IN1 | ((xor(xor(!(IN18), IN14 & IN27), !(IN36))) | IN6))))), IN2 & (IN1 | (xor(xor((!((!(IN15)) & IN33)) | ((xor(xor(!(IN47 & IN44), !(IN7 | IN29)), IN11)) | IN29), !(xor(xor((!(IN12 & IN39)) | false, (!(xor(xor(IN31, IN8), IN12))) & (!(xor(xor(IN28, IN6), IN10)))), (!(IN24 & IN26)) & IN19))), (IN13 & (!(xor(xor(IN49 | IN17, xor(xor(IN33, IN42), IN4)), !(IN24))))) | (xor(xor(xor(xor((!(IN50)) | (xor(xor(IN3, IN9), IN8)), IN37), IN19 | (xor(xor(IN12, IN20), IN44))), (IN33 & (IN26 & IN37)) & false), xor(xor((IN32 | IN14) & (IN48 | IN15), !(IN4)), !(IN3 | IN8)))))))), xor(xor(!((!(IN34)) | (((xor(xor((!(IN25)) & (!(IN43)), (IN23 | IN23) | (IN42 & IN28)), xor(xor(!(IN5), IN21 | IN11), IN50 & IN21))) & ((xor(xor(IN37, !(IN2)), !(IN8))) | (!(false & IN28)))) & (IN29 & (!((xor(xor(IN20, IN26), IN43)) & (!(IN5))))))), true), !((!(xor(xor(!(!(IN28 & IN27)), (xor(xor(!(IN2), xor(xor(IN41, IN6), IN50)), IN12 | IN21)) & (!(IN3 | IN13))), IN49))) | (!(IN18))))), (xor(xor(((((xor(xor(IN22, xor(xor(xor(xor(IN37, IN31), IN43), IN27 & IN11), !(IN25))), (!(IN40)) | (!(IN2)))) | IN7) | (!((!(!(IN44))) & (!(IN8 & IN24))))) & (!(xor(xor(!((IN26 & IN1) & IN16), (xor(xor(IN41 & IN1, IN32 & IN4), !(IN18))) & (!(xor(xor(IN44, IN21), IN15)))), (IN23 | (!(IN34))) | ((!(IN17)) & (IN46 & IN20)))))) | (IN41 | ((!((!(IN2 & IN40)) | (xor(xor(IN46 | IN27, IN36 | IN6), IN32 | IN27)))) & (IN45 & IN16))), (xor(xor(!(xor(xor(xor(xor((IN20 | IN41) & (xor(xor(IN5, IN20), IN39)), xor(xor(xor(xor(IN37, IN31), IN10), IN16 | IN46), IN23)), !(IN17)), IN24), ((xor(xor(IN17, IN3), IN42)) & (xor(xor(false, IN16), IN39))) | (xor(xor(IN3 & IN19, xor(xor(IN41, IN14), IN47)), IN34)))), IN24 | (!(IN14))), !(!(xor(xor(xor(xor(IN14 | IN36, xor(xor(IN23, IN17), IN46)), xor(xor(IN43, IN17), IN26)), (IN46 | IN37) & IN46), (xor(xor(IN8, IN26), IN43)) | (xor(xor(IN40, IN26), IN13))))))) & (xor(xor(IN19, IN10), IN40))), xor(xor(xor(xor((!(xor(xor((!(IN23)) & (!(IN4)), (xor(xor(IN26, IN41), IN36)) & (!(IN40))), (IN30 & IN42) & (IN34 | IN28)))) | (((!(IN26 & IN27)) & IN21) | IN10), IN31), IN33), IN45), ((!(IN15)) | ((IN11 & (!(IN41))) | ((xor(xor(IN38 & IN2, xor(xor(IN15, IN9), false)), !(IN31))) & ((IN3 | IN41) | (IN37 | IN31))))) & (!((((IN22 & IN49) & (xor(xor(IN49, IN14), IN33))) & (!(IN19 & IN10))) & IN43))))) & (!(IN50))), !((xor(xor(xor(xor(((xor(xor((IN29 | true) | IN10, xor(xor(xor(xor(IN46, IN7), IN5), IN26 & IN16), IN12)), (!(IN43)) | true)) | IN5) | (xor(xor(xor(xor((IN6 & IN18) & (IN49 & IN8), IN5 | (IN39 & IN35)), !(!(IN46))), ((xor(xor(IN10, IN40), IN6)) | (!(IN21))) & ((xor(xor(IN34, IN25), IN41)) & IN41)), IN33 | ((IN36 | true) & (IN12 & IN4)))), xor(xor(((xor(xor(IN12 | IN37, IN19), xor(xor(IN48, IN36), IN11))) | (xor(xor(IN34 | IN24, xor(xor(IN43, IN29), IN46)), xor(xor(IN9, IN7), IN3)))) | (((!(IN46)) & (xor(xor(IN41, IN21), IN12))) & IN43), IN15 | (!((!(IN15)) | (!(IN27))))), IN50)), (IN45 & (xor(xor(!(IN1), IN10), (!(IN12)) & (!(IN15))))) & (!(!(!(xor(xor(IN34, IN4), IN32)))))), (!((!(!(!(IN19)))) | (((xor(xor(IN49, IN25), IN23)) | (IN41 | IN31)) | (IN18 | (xor(xor(IN6, IN49), IN46)))))) | ((xor(xor(IN25, (!(IN6 | IN43)) | ((IN36 & IN19) & true)), false | IN41)) | IN37)), (!(((IN45 | (xor(xor(IN26, IN35), IN22))) | (xor(xor(IN20 & IN12, IN41 | IN12), IN20))) & (((IN38 & IN32) & (IN28 | IN14)) & (!(IN49 & IN15))))) | ((!((xor(xor(true & IN12, xor(xor(IN3, IN2), IN3)), IN20)) & (xor(xor(IN31, IN49), xor(xor(true, IN45), IN9))))) | (xor(xor((xor(xor(IN34 | IN2, IN13), xor(xor(IN34, IN10), IN43))) & IN49, ((xor(xor(IN4, IN7), IN45)) & IN6) | IN12), !(IN49 & (IN37 & IN8))))))) & (xor(xor(IN27, ((xor(xor(xor(xor((!(IN33)) | IN34, xor(xor(IN43 & IN37, xor(xor(IN25, IN31), IN29)), !(IN35))), (!(IN44)) | (IN36 | IN18)), IN10), !(IN23))) | ((xor(xor(!(IN13), IN36 | (true | IN25)), !(IN23 | IN16))) & (!(IN30)))) | (((xor(xor((IN43 & IN35) & IN36, !(!(IN2))), (!(IN13)) | IN30)) | ((!(IN2 | IN30)) & (xor(xor(xor(xor(IN3, IN17), IN29), IN45 | IN8), xor(xor(IN13, IN49), IN16))))) & ((xor(xor(xor(xor(IN28, IN25 | true), IN27), xor(xor(!(IN33), IN45 & IN24), !(IN6))), IN47)) | (!((xor(xor(IN6, IN25), IN24)) | (IN44 | IN22)))))), !(((xor(xor((false & IN49) & (xor(xor(IN16, IN18), IN50)), (!(IN23)) & (xor(xor(IN34, IN20), IN44))), (IN8 | IN3) & (!(IN32)))) | ((xor(xor(!(IN44), true & IN49), IN49)) | (IN15 | (xor(xor(IN5, IN32), IN2))))) & ((xor(xor(IN13 | (xor(xor(IN13, IN1), IN44)), (xor(xor(IN43, IN28), IN15)) | (xor(xor(IN21, IN37), IN45))), !(IN34 & IN2))) | (((IN34 & IN32) | IN29) & (!(xor(xor(IN18, IN4), IN40))))))))))

*)

FUNCTION_BLOCK F_CollectInput
  VAR_IN_OUT
      Data : ARRAY[1..50] OF BOOL;
  END_VAR
  VAR_INPUT
      TICK  : BOOL := 0;
      IN1   : BOOL := 0;
      IN2   : BOOL := 0;
      IN3   : BOOL := 0;
      IN4   : BOOL := 0;
      IN5   : BOOL := 0;
      RESET : BOOL := FALSE;
  END_VAR
  VAR_OUTPUT
      Finished : BOOL;
  END_VAR
  VAR
      j    : USINT := 1;
      tock : BOOL  := 0;
  END_VAR
  IF NOT RESET AND tock = NOT TICK THEN
      Data[j]   := IN1;
      Data[j+1] := IN2;
      Data[j+2] := IN3;
      Data[j+3] := IN4;
      Data[j+4] := IN5;
      j := j + 5;
      tock := TICK;
  ELSE
      j := 1;
      tock := 0;
  END_IF;
  Finished := (j > 50);
END_FUNCTION_BLOCK

PROGRAM Boiler
  VAR
    Data  : ARRAY[1..50] OF BOOL;
    Ready : BOOL;
    CollectInput : F_CollectInput;
  END_VAR
  VAR
    TICK     AT %IX1.0 : BOOL;
    IN1      AT %IX0.3 : BOOL;
    IN2      AT %IX0.4 : BOOL;
    IN3      AT %IX0.5 : BOOL;
    IN4      AT %IX0.6 : BOOL;
    IN5      AT %IX0.7 : BOOL;
    OutReady AT %QX0.0 : BOOL := FALSE;
    FeedNext AT %QX0.1 : BOOL := FALSE;
    Out      AT %QX0.2 : BOOL;
  END_VAR
  CollectInput(TICK:=TICK, IN1:=IN1, IN2:=IN2, IN3:=IN3, IN4:=IN4, IN5:=IN5);
  Ready := CollectInput.Finished;
  FeedNext := 1;
  IF Ready THEN
    Out := (((((NOT ((Data[45] XOR ((((((((Data[19] AND Data[49]) XOR (Data[3] AND Data[10])) XOR (NOT Data[13])) OR Data[18]) AND (Data[2] OR (((Data[32] XOR Data[39]) XOR Data[18]) OR Data[26]))) OR (NOT (((Data[23] AND Data[4]) AND (NOT Data[25])) AND (((NOT Data[15]) XOR ((Data[16] XOR Data[30]) XOR Data[44])) XOR ((Data[26] XOR TRUE) XOR Data[50]))))) XOR (NOT (((NOT ((Data[16] XOR Data[38]) XOR Data[11])) OR (Data[17] OR (NOT Data[22]))) OR (NOT (NOT (NOT Data[31])))))) XOR ((((NOT Data[2]) AND (NOT (Data[49] OR Data[20]))) AND (((Data[27] AND ((Data[47] XOR Data[2]) XOR TRUE)) XOR ((Data[21] OR Data[9]) OR Data[35])) XOR (Data[15] OR (NOT Data[16])))) AND ((NOT (NOT (NOT Data[17]))) OR (NOT ((Data[48] XOR (Data[15] AND Data[19])) XOR ((Data[13] XOR Data[36]) XOR Data[25]))))))) XOR (((Data[14] AND ((((((Data[38] AND Data[38]) AND (Data[45] OR Data[6])) XOR ((Data[12] AND Data[4]) OR (Data[47] OR Data[26]))) XOR ((((Data[2] XOR Data[1]) XOR Data[42]) XOR (Data[41] OR Data[2])) XOR (Data[43] OR Data[10]))) XOR ((NOT (Data[24] OR Data[39])) AND (((Data[35] OR Data[36]) XOR ((Data[4] XOR Data[46]) XOR Data[47])) XOR Data[50]))) XOR ((NOT ((Data[28] XOR Data[30]) XOR Data[39])) AND (((Data[49] XOR FALSE) XOR Data[31]) AND (Data[28] OR Data[47]))))) XOR Data[15]) XOR (NOT (Data[1] OR ((((NOT Data[18]) XOR (Data[14] AND Data[27])) XOR (NOT Data[36])) OR Data[6])))))) XOR (Data[2] AND (Data[1] OR ((((NOT ((NOT Data[15]) AND Data[33])) OR ((((NOT (Data[47] AND Data[44])) XOR (NOT (Data[7] OR Data[29]))) XOR Data[11]) OR Data[29])) XOR (NOT ((((NOT (Data[12] AND Data[39])) OR FALSE) XOR ((NOT ((Data[31] XOR Data[8]) XOR Data[12])) AND (NOT ((Data[28] XOR Data[6]) XOR Data[10])))) XOR ((NOT (Data[24] AND Data[26])) AND Data[19])))) XOR ((Data[13] AND (NOT (((Data[49] OR Data[17]) XOR ((Data[33] XOR Data[42]) XOR Data[4])) XOR (NOT Data[24])))) OR ((((((NOT Data[50]) OR ((Data[3] XOR Data[9]) XOR Data[8])) XOR Data[37]) XOR (Data[19] OR ((Data[12] XOR Data[20]) XOR Data[44]))) XOR ((Data[33] AND (Data[26] AND Data[37])) AND FALSE)) XOR ((((Data[32] OR Data[14]) AND (Data[48] OR Data[15])) XOR (NOT Data[4])) XOR (NOT (Data[3] OR Data[8]))))))))) XOR (((NOT ((NOT Data[34]) OR ((((((NOT Data[25]) AND (NOT Data[43])) XOR ((Data[23] OR Data[23]) OR (Data[42] AND Data[28]))) XOR (((NOT Data[5]) XOR (Data[21] OR Data[11])) XOR (Data[50] AND Data[21]))) AND (((Data[37] XOR (NOT Data[2])) XOR (NOT Data[8])) OR (NOT (FALSE AND Data[28])))) AND (Data[29] AND (NOT (((Data[20] XOR Data[26]) XOR Data[43]) AND (NOT Data[5]))))))) XOR TRUE) XOR (NOT ((NOT (((NOT (NOT (Data[28] AND Data[27]))) XOR ((((NOT Data[2]) XOR ((Data[41] XOR Data[6]) XOR Data[50])) XOR (Data[12] OR Data[21])) AND (NOT (Data[3] OR Data[13])))) XOR Data[49])) OR (NOT Data[18]))))) XOR (((((((((Data[22] XOR ((((Data[37] XOR Data[31]) XOR Data[43]) XOR (Data[27] AND Data[11])) XOR (NOT Data[25]))) XOR ((NOT Data[40]) OR (NOT Data[2]))) OR Data[7]) OR (NOT ((NOT (NOT Data[44])) AND (NOT (Data[8] AND Data[24]))))) AND (NOT (((NOT ((Data[26] AND Data[1]) AND Data[16])) XOR ((((Data[41] AND Data[1]) XOR (Data[32] AND Data[4])) XOR (NOT Data[18])) AND (NOT ((Data[44] XOR Data[21]) XOR Data[15])))) XOR ((Data[23] OR (NOT Data[34])) OR ((NOT Data[17]) AND (Data[46] AND Data[20])))))) OR (Data[41] OR ((NOT ((NOT (Data[2] AND Data[40])) OR (((Data[46] OR Data[27]) XOR (Data[36] OR Data[6])) XOR (Data[32] OR Data[27])))) AND (Data[45] AND Data[16])))) XOR ((((NOT ((((((Data[20] OR Data[41]) AND ((Data[5] XOR Data[20]) XOR Data[39])) XOR ((((Data[37] XOR Data[31]) XOR Data[10]) XOR (Data[16] OR Data[46])) XOR Data[23])) XOR (NOT Data[17])) XOR Data[24]) XOR ((((Data[17] XOR Data[3]) XOR Data[42]) AND ((FALSE XOR Data[16]) XOR Data[39])) OR (((Data[3] AND Data[19]) XOR ((Data[41] XOR Data[14]) XOR Data[47])) XOR Data[34])))) XOR (Data[24] OR (NOT Data[14]))) XOR (NOT (NOT (((((Data[14] OR Data[36]) XOR ((Data[23] XOR Data[17]) XOR Data[46])) XOR ((Data[43] XOR Data[17]) XOR Data[26])) XOR ((Data[46] OR Data[37]) AND Data[46])) XOR (((Data[8] XOR Data[26]) XOR Data[43]) OR ((Data[40] XOR Data[26]) XOR Data[13])))))) AND ((Data[19] XOR Data[10]) XOR Data[40]))) XOR ((((((NOT ((((NOT Data[23]) AND (NOT Data[4])) XOR (((Data[26] XOR Data[41]) XOR Data[36]) AND (NOT Data[40]))) XOR ((Data[30] AND Data[42]) AND (Data[34] OR Data[28])))) OR (((NOT (Data[26] AND Data[27])) AND Data[21]) OR Data[10])) XOR Data[31]) XOR Data[33]) XOR Data[45]) XOR (((NOT Data[15]) OR ((Data[11] AND (NOT Data[41])) OR ((((Data[38] AND Data[2]) XOR ((Data[15] XOR Data[9]) XOR FALSE)) XOR (NOT Data[31])) AND ((Data[3] OR Data[41]) OR (Data[37] OR Data[31]))))) AND (NOT ((((Data[22] AND Data[49]) AND ((Data[49] XOR Data[14]) XOR Data[33])) AND (NOT (Data[19] AND Data[10]))) AND Data[43]))))) AND (NOT Data[50]))) XOR (NOT (((((((((((Data[29] OR TRUE) OR Data[10]) XOR ((((Data[46] XOR Data[7]) XOR Data[5]) XOR (Data[26] AND Data[16])) XOR Data[12])) XOR ((NOT Data[43]) OR TRUE)) OR Data[5]) OR ((((((Data[6] AND Data[18]) AND (Data[49] AND Data[8])) XOR (Data[5] OR (Data[39] AND Data[35]))) XOR (NOT (NOT Data[46]))) XOR ((((Data[10] XOR Data[40]) XOR Data[6]) OR (NOT Data[21])) AND (((Data[34] XOR Data[25]) XOR Data[41]) AND Data[41]))) XOR (Data[33] OR ((Data[36] OR TRUE) AND (Data[12] AND Data[4]))))) XOR (((((((Data[12] OR Data[37]) XOR Data[19]) XOR ((Data[48] XOR Data[36]) XOR Data[11])) OR (((Data[34] OR Data[24]) XOR ((Data[43] XOR Data[29]) XOR Data[46])) XOR ((Data[9] XOR Data[7]) XOR Data[3]))) OR (((NOT Data[46]) AND ((Data[41] XOR Data[21]) XOR Data[12])) AND Data[43])) XOR (Data[15] OR (NOT ((NOT Data[15]) OR (NOT Data[27]))))) XOR Data[50])) XOR ((Data[45] AND (((NOT Data[1]) XOR Data[10]) XOR ((NOT Data[12]) AND (NOT Data[15])))) AND (NOT (NOT (NOT ((Data[34] XOR Data[4]) XOR Data[32])))))) XOR ((NOT ((NOT (NOT (NOT Data[19]))) OR ((((Data[49] XOR Data[25]) XOR Data[23]) OR (Data[41] OR Data[31])) OR (Data[18] OR ((Data[6] XOR Data[49]) XOR Data[46]))))) OR (((Data[25] XOR ((NOT (Data[6] OR Data[43])) OR ((Data[36] AND Data[19]) AND TRUE))) XOR (FALSE OR Data[41])) OR Data[37]))) XOR ((NOT (((Data[45] OR ((Data[26] XOR Data[35]) XOR Data[22])) OR (((Data[20] AND Data[12]) XOR (Data[41] OR Data[12])) XOR Data[20])) AND (((Data[38] AND Data[32]) AND (Data[28] OR Data[14])) AND (NOT (Data[49] AND Data[15]))))) OR ((NOT ((((TRUE AND Data[12]) XOR ((Data[3] XOR Data[2]) XOR Data[3])) XOR Data[20]) AND ((Data[31] XOR Data[49]) XOR ((TRUE XOR Data[45]) XOR Data[9])))) OR ((((((Data[34] OR Data[2]) XOR Data[13]) XOR ((Data[34] XOR Data[10]) XOR Data[43])) AND Data[49]) XOR ((((Data[4] XOR Data[7]) XOR Data[45]) AND Data[6]) OR Data[12])) XOR (NOT (Data[49] AND (Data[37] AND Data[8]))))))) AND ((Data[27] XOR ((((((((NOT Data[33]) OR Data[34]) XOR (((Data[43] AND Data[37]) XOR ((Data[25] XOR Data[31]) XOR Data[29])) XOR (NOT Data[35]))) XOR ((NOT Data[44]) OR (Data[36] OR Data[18]))) XOR Data[10]) XOR (NOT Data[23])) OR ((((NOT Data[13]) XOR (Data[36] OR (TRUE OR Data[25]))) XOR (NOT (Data[23] OR Data[16]))) AND (NOT Data[30]))) OR ((((((Data[43] AND Data[35]) AND Data[36]) XOR (NOT (NOT Data[2]))) XOR ((NOT Data[13]) OR Data[30])) OR ((NOT (Data[2] OR Data[30])) AND ((((Data[3] XOR Data[17]) XOR Data[29]) XOR (Data[45] OR Data[8])) XOR ((Data[13] XOR Data[49]) XOR Data[16])))) AND (((((Data[28] XOR (Data[25] OR TRUE)) XOR Data[27]) XOR (((NOT Data[33]) XOR (Data[45] AND Data[24])) XOR (NOT Data[6]))) XOR Data[47]) OR (NOT (((Data[6] XOR Data[25]) XOR Data[24]) OR (Data[44] OR Data[22]))))))) XOR (NOT ((((((FALSE AND Data[49]) AND ((Data[16] XOR Data[18]) XOR Data[50])) XOR ((NOT Data[23]) AND ((Data[34] XOR Data[20]) XOR Data[44]))) XOR ((Data[8] OR Data[3]) AND (NOT Data[32]))) OR ((((NOT Data[44]) XOR (TRUE AND Data[49])) XOR Data[49]) OR (Data[15] OR ((Data[5] XOR Data[32]) XOR Data[2])))) AND ((((Data[13] OR ((Data[13] XOR Data[1]) XOR Data[44])) XOR (((Data[43] XOR Data[28]) XOR Data[15]) OR ((Data[21] XOR Data[37]) XOR Data[45]))) XOR (NOT (Data[34] AND Data[2]))) OR (((Data[34] AND Data[32]) OR Data[29]) AND (NOT ((Data[18] XOR Data[4]) XOR Data[40]))))))))));
    OutReady := 1;
    CollectInput(RESET:=TRUE);
  END_IF;
END_PROGRAM

CONFIGURATION Config0
  RESOURCE Res0 ON PLC
    TASK task0(INTERVAL := T#20ms,PRIORITY := 0);
    PROGRAM instance0 WITH task0 : Boiler;
  END_RESOURCE
END_CONFIGURATION

(* ---- RND-EXPR_folky-amigo-bails.st ---- *)
(*
This code implements a randomly grown symbolic expression:

(xor(xor(IN49, xor(xor(xor(xor(xor(xor(((!(xor(xor(IN40, IN39), IN45))) & (((IN22 | IN24) & IN8) | (!(false | IN1)))) | (IN15 | (((!(IN10)) & (IN37 | IN3)) | (!(xor(xor(IN33, IN28), IN50))))), (xor(xor(IN22, IN43 | (!(IN15 & IN23))), (xor(xor(!(IN37), true), xor(xor(IN39, IN32), IN13))) & IN50)) & (!((xor(xor(xor(xor(IN14, IN18), IN6), IN41), IN34)) | (xor(xor(!(IN42), IN41), IN50 & IN1))))), !(xor(xor(!(xor(xor(xor(xor(IN1, IN30), IN23), IN23 & IN2), !(IN27))), !(!(IN37 | IN35))), ((IN16 & IN7) & (xor(xor(IN49, IN41), IN17))) & (!(!(IN16)))))), (((xor(xor((IN9 & IN49) | (xor(xor(IN37, IN18), IN18)), xor(xor(!(IN25), !(IN7)), IN30)), !(IN37 & IN40))) & (!(IN23))) & ((!(!(!(IN43)))) | (IN21 | (xor(xor(IN12 | IN36, IN43 | IN1), IN42 | IN13))))) | (((xor(xor(IN31, (xor(true, IN22)) & (IN32 | IN17)), IN46)) | (((true | IN47) | (xor(xor(IN5, IN43), IN31))) | (xor(xor(IN16 & IN37, !(IN42)), !(IN46))))) | IN36)), IN23), xor(xor(xor(xor(IN4, IN48), IN22), (xor(xor(((!(IN44 | IN31)) & (!(IN47 & IN36))) | ((!(IN25)) & (xor(xor(IN28 & IN45, IN48 & IN43), IN33))), (!(!(IN27 | IN28))) | (!(xor(xor(!(IN3), IN37 | IN22), xor(xor(IN47, true), IN44))))), !(!(xor(xor(IN34 | IN7, !(IN8)), xor(xor(IN22, IN12), IN27)))))) & ((xor(xor((IN23 & (!(IN36))) | ((IN38 | IN39) | (IN28 & IN38)), (!(IN1)) | IN33), ((IN12 & IN8) | (IN40 | IN33)) & (IN20 | (IN12 | IN35)))) & (!(((xor(xor(IN26, IN19), IN21)) | IN43) | (!(xor(xor(IN18, IN27), IN47))))))), IN22)), xor(xor(xor(xor(!(IN38), (!(xor(xor((IN45 | IN28) | (xor(xor(IN10, IN30), IN29)), xor(xor(!(IN49), xor(xor(IN29, IN34), IN2)), IN34)), (!(IN39)) | (xor(xor(IN26, IN43), IN12))))) | IN33), (!(((!(IN16)) | (IN37 & IN45)) | ((IN29 & IN31) & IN41))) | (xor(xor(!(xor(xor(IN30 & IN10, xor(xor(IN1, IN15), IN6)), true)), xor(xor((xor(xor(IN45, IN15), IN38)) & (IN8 & IN42), !(IN18 | IN39)), IN46)), !((!(IN36)) & (!(IN9)))))), xor(xor(!((xor(xor(xor(xor(!(IN9), xor(xor(IN24, IN25), IN12)), xor(xor(IN50, IN31), IN45)), (IN34 | IN22) & (IN8 & IN18)), (xor(xor(IN7, IN2), IN36)) & (xor(xor(IN12, IN41), IN20)))) & (!(!(IN41 & IN39)))), xor(xor(!((xor(xor(!(IN20), IN27 & IN35), xor(xor(IN43, IN36), IN10))) | IN37), (xor(xor(!(IN25 & IN21), (xor(xor(IN26, IN27), IN8)) | (IN2 | IN17)), (!(IN3)) & (!(IN33)))) & ((xor(xor(xor(xor(IN2, IN27), IN8), !(IN39)), IN10)) | IN47)), xor(xor(!((IN46 | IN24) & (IN18 & IN45)), IN36), xor(xor(IN16, !(xor(xor(IN26, IN5), IN21))), !(IN18 | IN25))))), IN50)), (xor(xor(IN13, IN40), xor(xor(xor(xor(xor(xor(true | IN46, IN7 | IN15), IN23 & IN31), (xor(xor(IN44, IN27), IN22)) & (IN30 | IN22)), (IN3 & IN38) | IN26), xor(xor(IN47, xor(xor(!(IN28), xor(xor(IN47, IN7), IN1)), IN49)), xor(xor(!(IN47), IN19 | IN47), IN33))), !(!(!(IN27)))))) | (xor(xor(IN26, xor(xor(!(!(IN14)), !(IN11)), (IN22 & (IN1 & IN37)) & IN45)), IN22))))), !((!(xor(xor((xor(xor((IN33 | IN35) & (IN23 & IN20), (xor(xor(IN37, IN42), IN41)) | (IN10 | IN41)), xor(xor(xor(xor(IN48, IN43), IN20), xor(xor(false, IN26), IN33)), !(IN7)))) & (((IN24 | IN23) & (IN13 & IN2)) | ((IN7 | IN31) & (IN16 & IN26))), (!(!(xor(xor(IN20, IN20), IN27)))) | ((xor(xor(IN39 | IN18, IN48 & IN19), IN26 | IN50)) | (!(IN21 & true)))), IN35))) | ((xor(xor(IN3, xor(xor(!(IN28 & (IN36 & IN20)), !(!(IN8 | IN18))), IN7)), (IN29 & ((IN47 | IN26) & (IN34 | IN39))) | ((IN31 | (xor(xor(IN13, IN20), IN41))) & (!(!(IN4)))))) & (!(xor(xor((!(!(IN25))) & (!(xor(xor(IN37, IN37), IN2))), (!(xor(xor(IN6, IN5), IN39))) & (IN30 | (!(IN36)))), (IN4 & (!(IN36))) & (IN45 | (!(IN11)))))))))) & ((xor(xor(xor(xor(xor(xor(IN27, (((!(IN4)) | ((IN18 & IN27) & IN1)) & IN18) | IN11), !(xor(xor(IN50, xor(xor(xor(xor(!(IN47), !(IN15)), xor(xor(IN22, IN6), IN39)), xor(xor(!(IN7), xor(xor(IN20, IN45), IN23)), IN11 | IN44)), (xor(xor(IN35, IN30), IN47)) & IN21)), ((IN46 & IN40) & (!(IN42))) & ((IN11 | IN48) | IN50)))), !(xor(xor(!(IN3), (!((IN6 & IN14) & (!(IN48)))) & ((xor(xor(IN11 | IN32, IN37 & IN43), xor(xor(IN14, IN46), IN46))) & (xor(xor(IN13 & IN1, IN6), IN26 & IN2)))), IN15 & (((!(IN42)) & (IN17 | true)) & (xor(xor(xor(xor(IN18, true), IN38), IN28), IN5 | IN48)))))), ((xor(xor(!(xor(xor(xor(xor(true, IN21), IN4), IN5 | IN29), xor(xor(IN14, IN8), IN32))), xor(xor(!(IN39 & IN46), (!(IN23)) | IN6), xor(xor(xor(xor(IN4, IN7), IN39), IN42), xor(xor(IN24, IN27), IN13)))), IN32)) | (!(!((IN20 & IN42) & (IN32 & IN34))))) | (!(((xor(xor(IN20 & IN9, IN41 | IN22), IN39 | IN1)) | (!(IN10 | true))) & IN33))), xor(xor(((((IN34 & (IN34 | IN19)) & (xor(xor(!(IN38), IN16 & false), IN25 & IN42))) & (!(IN43 | (xor(xor(IN25, IN19), IN23))))) & (((xor(xor(xor(xor(IN19, IN47), IN29), !(IN40)), xor(xor(IN48, IN12), IN14))) | ((IN38 | IN34) | (!(IN32)))) & (((!(IN31)) | (IN31 | IN33)) | (!(IN26 | IN30))))) | ((IN50 & IN24) & (!(xor(xor(!(IN48), IN44), !(xor(xor(IN39, IN12), IN9)))))), IN4), xor(xor(((xor(xor(xor(xor(IN48 & IN33, !(IN27)), !(IN10)), IN3), xor(xor(IN23 & IN25, xor(xor(IN41, IN18), IN43)), IN29 & IN26))) & (xor(xor(xor(xor(xor(xor(IN29, IN43), IN9), xor(xor(false, IN36), IN30)), xor(xor(IN5, IN39), IN21)), !(xor(xor(IN12, IN45), IN39))), xor(xor(IN34 | IN22, IN33 | IN28), IN31 & IN41)))) | (((xor(xor(IN18 | IN1, xor(xor(IN48, IN49), IN30)), IN15)) & (xor(xor(IN5, IN10 & IN33), xor(xor(IN22, IN10), IN14)))) & (!((IN6 & IN13) & (!(IN7))))), (!((xor(xor(IN42 & IN45, IN13 | IN15), xor(xor(IN21, IN7), true))) | IN24)) & (xor(xor(((IN9 & IN10) & (IN46 | IN1)) | ((IN23 | IN33) & (!(IN24))), !((xor(xor(IN3, IN33), IN12)) & (true | IN46))), (xor(xor(IN43 & IN10, false & IN14), IN26 | IN41)) & ((IN44 | IN25) | (!(IN40)))))), !(xor(xor(IN31, !(IN46 & IN10)), (IN1 | (IN2 & IN8)) & (xor(xor(IN22, !(IN44)), false | IN11))))))), (IN1 & (xor(xor(IN15, (xor(xor(!(true & IN28), !(IN39)), IN31)) | (!(IN38 & IN44))), xor(xor(IN42 | IN35, xor(xor((IN31 & IN14) | (!(IN19)), (IN31 | IN38) & IN49), IN47 & (!(IN14)))), xor(xor(IN31 | (IN37 | IN24), IN1), !(IN44)))))) & (!(xor(xor((false | ((IN49 | IN21) | IN37)) & ((xor(xor(IN21 & IN40, IN6 & IN19), IN7 | IN21)) | (xor(xor(!(IN47), IN46 | IN49), IN33 & IN4))), !(!(!(xor(xor(IN30, IN24), IN17))))), ((!(IN46 | IN46)) | (!(!(IN41)))) & (!(xor(xor(IN24 | IN26, !(IN33)), IN21 & IN27)))))))) | IN24)

*)

FUNCTION_BLOCK F_CollectInput
  VAR_IN_OUT
      Data : ARRAY[1..50] OF BOOL;
  END_VAR
  VAR_INPUT
      TICK  : BOOL := 0;
      IN1   : BOOL := 0;
      IN2   : BOOL := 0;
      IN3   : BOOL := 0;
      IN4   : BOOL := 0;
      IN5   : BOOL := 0;
      RESET : BOOL := FALSE;
  END_VAR
  VAR_OUTPUT
      Finished : BOOL;
  END_VAR
  VAR
      j    : USINT := 1;
      tock : BOOL  := 0;
  END_VAR
  IF NOT RESET AND tock = NOT TICK THEN
      Data[j]   := IN1;
      Data[j+1] := IN2;
      Data[j+2] := IN3;
      Data[j+3] := IN4;
      Data[j+4] := IN5;
      j := j + 5;
      tock := TICK;
  ELSE
      j := 1;
      tock := 0;
  END_IF;
  Finished := (j > 50);
END_FUNCTION_BLOCK

PROGRAM Boiler
  VAR
    Data  : ARRAY[1..50] OF BOOL;
    Ready : BOOL;
    CollectInput : F_CollectInput;
  END_VAR
  VAR
    TICK     AT %IX1.0 : BOOL;
    IN1      AT %IX0.3 : BOOL;
    IN2      AT %IX0.4 : BOOL;
    IN3      AT %IX0.5 : BOOL;
    IN4      AT %IX0.6 : BOOL;
    IN5      AT %IX0.7 : BOOL;
    OutReady AT %QX0.0 : BOOL := FALSE;
    FeedNext AT %QX0.1 : BOOL := FALSE;
    Out      AT %QX0.2 : BOOL;
  END_VAR
  CollectInput(TICK:=TICK, IN1:=IN1, IN2:=IN2, IN3:=IN3, IN4:=IN4, IN5:=IN5);
  Ready := CollectInput.Finished;
  FeedNext := 1;
  IF Ready THEN
    Out := (((Data[49] XOR (((((((((NOT ((Data[40] XOR Data[39]) XOR Data[45])) AND (((Data[22] OR Data[24]) AND Data[8]) OR (NOT (FALSE OR Data[1])))) OR (Data[15] OR (((NOT Data[10]) AND (Data[37] OR Data[3])) OR (NOT ((Data[33] XOR Data[28]) XOR Data[50]))))) XOR (((Data[22] XOR (Data[43] OR (NOT (Data[15] AND Data[23])))) XOR ((((NOT Data[37]) XOR TRUE) XOR ((Data[39] XOR Data[32]) XOR Data[13])) AND Data[50])) AND (NOT (((((Data[14] XOR Data[18]) XOR Data[6]) XOR Data[41]) XOR Data[34]) OR (((NOT Data[42]) XOR Data[41]) XOR (Data[50] AND Data[1])))))) XOR (NOT (((NOT ((((Data[1] XOR Data[30]) XOR Data[23]) XOR (Data[23] AND Data[2])) XOR (NOT Data[27]))) XOR (NOT (NOT (Data[37] OR Data[35])))) XOR (((Data[16] AND Data[7]) AND ((Data[49] XOR Data[41]) XOR Data[17])) AND (NOT (NOT Data[16])))))) XOR (((((((Data[9] AND Data[49]) OR ((Data[37] XOR Data[18]) XOR Data[18])) XOR (((NOT Data[25]) XOR (NOT Data[7])) XOR Data[30])) XOR (NOT (Data[37] AND Data[40]))) AND (NOT Data[23])) AND ((NOT (NOT (NOT Data[43]))) OR (Data[21] OR (((Data[12] OR Data[36]) XOR (Data[43] OR Data[1])) XOR (Data[42] OR Data[13]))))) OR ((((Data[31] XOR ((TRUE XOR Data[22]) AND (Data[32] OR Data[17]))) XOR Data[46]) OR (((TRUE OR Data[47]) OR ((Data[5] XOR Data[43]) XOR Data[31])) OR (((Data[16] AND Data[37]) XOR (NOT Data[42])) XOR (NOT Data[46])))) OR Data[36]))) XOR Data[23]) XOR ((((Data[4] XOR Data[48]) XOR Data[22]) XOR ((((((NOT (Data[44] OR Data[31])) AND (NOT (Data[47] AND Data[36]))) OR ((NOT Data[25]) AND (((Data[28] AND Data[45]) XOR (Data[48] AND Data[43])) XOR Data[33]))) XOR ((NOT (NOT (Data[27] OR Data[28]))) OR (NOT (((NOT Data[3]) XOR (Data[37] OR Data[22])) XOR ((Data[47] XOR TRUE) XOR Data[44]))))) XOR (NOT (NOT (((Data[34] OR Data[7]) XOR (NOT Data[8])) XOR ((Data[22] XOR Data[12]) XOR Data[27]))))) AND (((((Data[23] AND (NOT Data[36])) OR ((Data[38] OR Data[39]) OR (Data[28] AND Data[38]))) XOR ((NOT Data[1]) OR Data[33])) XOR (((Data[12] AND Data[8]) OR (Data[40] OR Data[33])) AND (Data[20] OR (Data[12] OR Data[35])))) AND (NOT ((((Data[26] XOR Data[19]) XOR Data[21]) OR Data[43]) OR (NOT ((Data[18] XOR Data[27]) XOR Data[47]))))))) XOR Data[22])) XOR (((((NOT Data[38]) XOR ((NOT ((((Data[45] OR Data[28]) OR ((Data[10] XOR Data[30]) XOR Data[29])) XOR (((NOT Data[49]) XOR ((Data[29] XOR Data[34]) XOR Data[2])) XOR Data[34])) XOR ((NOT Data[39]) OR ((Data[26] XOR Data[43]) XOR Data[12])))) OR Data[33])) XOR ((NOT (((NOT Data[16]) OR (Data[37] AND Data[45])) OR ((Data[29] AND Data[31]) AND Data[41]))) OR (((NOT (((Data[30] AND Data[10]) XOR ((Data[1] XOR Data[15]) XOR Data[6])) XOR TRUE)) XOR (((((Data[45] XOR Data[15]) XOR Data[38]) AND (Data[8] AND Data[42])) XOR (NOT (Data[18] OR Data[39]))) XOR Data[46])) XOR (NOT ((NOT Data[36]) AND (NOT Data[9])))))) XOR (((NOT ((((((NOT Data[9]) XOR ((Data[24] XOR Data[25]) XOR Data[12])) XOR ((Data[50] XOR Data[31]) XOR Data[45])) XOR ((Data[34] OR Data[22]) AND (Data[8] AND Data[18]))) XOR (((Data[7] XOR Data[2]) XOR Data[36]) AND ((Data[12] XOR Data[41]) XOR Data[20]))) AND (NOT (NOT (Data[41] AND Data[39]))))) XOR (((NOT ((((NOT Data[20]) XOR (Data[27] AND Data[35])) XOR ((Data[43] XOR Data[36]) XOR Data[10])) OR Data[37])) XOR ((((NOT (Data[25] AND Data[21])) XOR (((Data[26] XOR Data[27]) XOR Data[8]) OR (Data[2] OR Data[17]))) XOR ((NOT Data[3]) AND (NOT Data[33]))) AND (((((Data[2] XOR Data[27]) XOR Data[8]) XOR (NOT Data[39])) XOR Data[10]) OR Data[47]))) XOR (((NOT ((Data[46] OR Data[24]) AND (Data[18] AND Data[45]))) XOR Data[36]) XOR ((Data[16] XOR (NOT ((Data[26] XOR Data[5]) XOR Data[21]))) XOR (NOT (Data[18] OR Data[25])))))) XOR Data[50])) XOR (((Data[13] XOR Data[40]) XOR (((((((TRUE OR Data[46]) XOR (Data[7] OR Data[15])) XOR (Data[23] AND Data[31])) XOR (((Data[44] XOR Data[27]) XOR Data[22]) AND (Data[30] OR Data[22]))) XOR ((Data[3] AND Data[38]) OR Data[26])) XOR ((Data[47] XOR (((NOT Data[28]) XOR ((Data[47] XOR Data[7]) XOR Data[1])) XOR Data[49])) XOR (((NOT Data[47]) XOR (Data[19] OR Data[47])) XOR Data[33]))) XOR (NOT (NOT (NOT Data[27]))))) OR ((Data[26] XOR (((NOT (NOT Data[14])) XOR (NOT Data[11])) XOR ((Data[22] AND (Data[1] AND Data[37])) AND Data[45]))) XOR Data[22]))))) XOR (NOT ((NOT (((((((Data[33] OR Data[35]) AND (Data[23] AND Data[20])) XOR (((Data[37] XOR Data[42]) XOR Data[41]) OR (Data[10] OR Data[41]))) XOR ((((Data[48] XOR Data[43]) XOR Data[20]) XOR ((FALSE XOR Data[26]) XOR Data[33])) XOR (NOT Data[7]))) AND (((Data[24] OR Data[23]) AND (Data[13] AND Data[2])) OR ((Data[7] OR Data[31]) AND (Data[16] AND Data[26])))) XOR ((NOT (NOT ((Data[20] XOR Data[20]) XOR Data[27]))) OR ((((Data[39] OR Data[18]) XOR (Data[48] AND Data[19])) XOR (Data[26] OR Data[50])) OR (NOT (Data[21] AND TRUE))))) XOR Data[35])) OR (((Data[3] XOR (((NOT (Data[28] AND (Data[36] AND Data[20]))) XOR (NOT (NOT (Data[8] OR Data[18])))) XOR Data[7])) XOR ((Data[29] AND ((Data[47] OR Data[26]) AND (Data[34] OR Data[39]))) OR ((Data[31] OR ((Data[13] XOR Data[20]) XOR Data[41])) AND (NOT (NOT Data[4]))))) AND (NOT ((((NOT (NOT Data[25])) AND (NOT ((Data[37] XOR Data[37]) XOR Data[2]))) XOR ((NOT ((Data[6] XOR Data[5]) XOR Data[39])) AND (Data[30] OR (NOT Data[36])))) XOR ((Data[4] AND (NOT Data[36])) AND (Data[45] OR (NOT Data[11]))))))))) AND (((((((Data[27] XOR ((((NOT Data[4]) OR ((Data[18] AND Data[27]) AND Data[1])) AND Data[18]) OR Data[11])) XOR (NOT ((Data[50] XOR (((((NOT Data[47]) XOR (NOT Data[15])) XOR ((Data[22] XOR Data[6]) XOR Data[39])) XOR (((NOT Data[7]) XOR ((Data[20] XOR Data[45]) XOR Data[23])) XOR (Data[11] OR Data[44]))) XOR (((Data[35] XOR Data[30]) XOR Data[47]) AND Data[21]))) XOR (((Data[46] AND Data[40]) AND (NOT Data[42])) AND ((Data[11] OR Data[48]) OR Data[50]))))) XOR (NOT (((NOT Data[3]) XOR ((NOT ((Data[6] AND Data[14]) AND (NOT Data[48]))) AND ((((Data[11] OR Data[32]) XOR (Data[37] AND Data[43])) XOR ((Data[14] XOR Data[46]) XOR Data[46])) AND (((Data[13] AND Data[1]) XOR Data[6]) XOR (Data[26] AND Data[2]))))) XOR (Data[15] AND (((NOT Data[42]) AND (Data[17] OR TRUE)) AND ((((Data[18] XOR TRUE) XOR Data[38]) XOR Data[28]) XOR (Data[5] OR Data[48]))))))) XOR (((((NOT ((((TRUE XOR Data[21]) XOR Data[4]) XOR (Data[5] OR Data[29])) XOR ((Data[14] XOR Data[8]) XOR Data[32]))) XOR (((NOT (Data[39] AND Data[46])) XOR ((NOT Data[23]) OR Data[6])) XOR ((((Data[4] XOR Data[7]) XOR Data[39]) XOR Data[42]) XOR ((Data[24] XOR Data[27]) XOR Data[13])))) XOR Data[32]) OR (NOT (NOT ((Data[20] AND Data[42]) AND (Data[32] AND Data[34]))))) OR (NOT (((((Data[20] AND Data[9]) XOR (Data[41] OR Data[22])) XOR (Data[39] OR Data[1])) OR (NOT (Data[10] OR TRUE))) AND Data[33])))) XOR (((((((Data[34] AND (Data[34] OR Data[19])) AND (((NOT Data[38]) XOR (Data[16] AND FALSE)) XOR (Data[25] AND Data[42]))) AND (NOT (Data[43] OR ((Data[25] XOR Data[19]) XOR Data[23])))) AND ((((((Data[19] XOR Data[47]) XOR Data[29]) XOR (NOT Data[40])) XOR ((Data[48] XOR Data[12]) XOR Data[14])) OR ((Data[38] OR Data[34]) OR (NOT Data[32]))) AND (((NOT Data[31]) OR (Data[31] OR Data[33])) OR (NOT (Data[26] OR Data[30]))))) OR ((Data[50] AND Data[24]) AND (NOT (((NOT Data[48]) XOR Data[44]) XOR (NOT ((Data[39] XOR Data[12]) XOR Data[9])))))) XOR Data[4]) XOR (((((((((Data[48] AND Data[33]) XOR (NOT Data[27])) XOR (NOT Data[10])) XOR Data[3]) XOR (((Data[23] AND Data[25]) XOR ((Data[41] XOR Data[18]) XOR Data[43])) XOR (Data[29] AND Data[26]))) AND ((((((Data[29] XOR Data[43]) XOR Data[9]) XOR ((FALSE XOR Data[36]) XOR Data[30])) XOR ((Data[5] XOR Data[39]) XOR Data[21])) XOR (NOT ((Data[12] XOR Data[45]) XOR Data[39]))) XOR (((Data[34] OR Data[22]) XOR (Data[33] OR Data[28])) XOR (Data[31] AND Data[41])))) OR (((((Data[18] OR Data[1]) XOR ((Data[48] XOR Data[49]) XOR Data[30])) XOR Data[15]) AND ((Data[5] XOR (Data[10] AND Data[33])) XOR ((Data[22] XOR Data[10]) XOR Data[14]))) AND (NOT ((Data[6] AND Data[13]) AND (NOT Data[7]))))) XOR ((NOT ((((Data[42] AND Data[45]) XOR (Data[13] OR Data[15])) XOR ((Data[21] XOR Data[7]) XOR TRUE)) OR Data[24])) AND (((((Data[9] AND Data[10]) AND (Data[46] OR Data[1])) OR ((Data[23] OR Data[33]) AND (NOT Data[24]))) XOR (NOT (((Data[3] XOR Data[33]) XOR Data[12]) AND (TRUE OR Data[46])))) XOR ((((Data[43] AND Data[10]) XOR (FALSE AND Data[14])) XOR (Data[26] OR Data[41])) AND ((Data[44] OR Data[25]) OR (NOT Data[40])))))) XOR (NOT ((Data[31] XOR (NOT (Data[46] AND Data[10]))) XOR ((Data[1] OR (Data[2] AND Data[8])) AND ((Data[22] XOR (NOT Data[44])) XOR (FALSE OR Data[11])))))))) XOR ((Data[1] AND ((Data[15] XOR ((((NOT (TRUE AND Data[28])) XOR (NOT Data[39])) XOR Data[31]) OR (NOT (Data[38] AND Data[44])))) XOR (((Data[42] OR Data[35]) XOR ((((Data[31] AND Data[14]) OR (NOT Data[19])) XOR ((Data[31] OR Data[38]) AND Data[49])) XOR (Data[47] AND (NOT Data[14])))) XOR (((Data[31] OR (Data[37] OR Data[24])) XOR Data[1]) XOR (NOT Data[44]))))) AND (NOT ((((FALSE OR ((Data[49] OR Data[21]) OR Data[37])) AND ((((Data[21] AND Data[40]) XOR (Data[6] AND Data[19])) XOR (Data[7] OR Data[21])) OR (((NOT Data[47]) XOR (Data[46] OR Data[49])) XOR (Data[33] AND Data[4])))) XOR (NOT (NOT (NOT ((Data[30] XOR Data[24]) XOR Data[17]))))) XOR (((NOT (Data[46] OR Data[46])) OR (NOT (NOT Data[41]))) AND (NOT (((Data[24] OR Data[26]) XOR (NOT Data[33])) XOR (Data[21] AND Data[27])))))))) OR Data[24]));
    OutReady := 1;
    CollectInput(RESET:=TRUE);
  END_IF;
END_PROGRAM

CONFIGURATION Config0
  RESOURCE Res0 ON PLC
    TASK task0(INTERVAL := T#20ms,PRIORITY := 0);
    PROGRAM instance0 WITH task0 : Boiler;
  END_RESOURCE
END_CONFIGURATION

(* ---- RND-EXPR_holly-stave-heady.st ---- *)
(*
This code implements a randomly grown symbolic expression:

xor(xor(xor(xor(IN21, (IN18 & (xor(xor(((xor(xor((IN50 | IN1) & (IN14 & IN11), xor(xor(IN43 | IN14, xor(xor(IN44, IN33), IN13)), !(IN12))), IN23)) | (xor(xor((!(IN4)) & (!(IN36)), (IN18 | IN26) | (IN35 | IN4)), IN17))) | (IN48 | (!((xor(xor(IN18, IN37), IN11)) | IN15))), IN14 & (!(IN48))), IN43 & (xor(xor(xor(xor((!(IN37)) & (IN28 & IN40), IN2), (!(IN3)) | (IN40 & IN12)), xor(xor(xor(xor(IN28 & IN23, IN41), !(IN32)), (!(IN47)) & (!(IN32))), (!(IN12)) | (xor(xor(IN29, false), IN29)))), xor(xor(xor(xor(!(IN14), !(IN13)), IN21 | IN22), xor(xor(!(IN43), IN19 | IN33), xor(xor(IN36, IN14), IN24))), true)))))) & ((IN35 | IN16) | IN50)), xor(xor(IN42, IN33), IN47)), xor(xor(((!((xor(xor((IN10 | (xor(xor(IN36, IN36), IN48))) | ((!(IN42)) & (IN8 | IN31)), ((!(IN11)) | (IN12 & IN9)) | ((xor(xor(IN8, IN5), IN3)) | (true | IN26))), !((IN24 | IN50) & (xor(xor(IN15, IN45), IN38))))) & (xor(xor(IN42 | ((IN18 | IN37) & (IN15 & IN43)), (!(IN15)) | ((IN25 | IN45) | (xor(xor(IN19, IN35), IN4)))), IN3 | (!(IN13 | IN38)))))) | (IN14 | ((xor(xor(((!(IN1)) | (IN2 & IN27)) & ((IN45 | IN39) & false), xor(xor(!(!(IN21)), IN27), (IN19 | IN19) | (IN14 | IN32))), (xor(xor(xor(xor(true, IN5), IN21), xor(xor(IN38, IN6), IN18)), xor(xor(IN2, IN3), true))) & (!(IN44 & IN27)))) | (!(((IN5 & IN37) & IN1) | ((IN18 & IN28) & (IN33 | IN49))))))) | (!(!((!(IN26)) | (!((xor(xor(IN23 | IN42, !(IN8)), !(IN5))) & ((IN8 & IN13) & (xor(xor(IN36, IN2), IN28)))))))), (xor(xor(IN48, xor(xor(IN37 & (xor(xor(IN8, IN38), (!(IN20 | IN8)) | ((IN32 | IN43) & (!(IN9))))), (!(IN28 | (xor(xor(IN40 & IN12, !(IN46)), IN17 & IN49)))) | IN38), IN3)), xor(xor(!(!(xor(xor(xor(xor(!(IN23), IN1), IN18 & IN50), !(!(IN11))), xor(xor(xor(xor(IN47, IN15), IN49), !(IN44)), !(IN44))))), xor(xor(xor(xor((!(IN29 | IN44)) | IN43, IN34), xor(xor(xor(xor(IN8 & IN46, IN14), IN25 & IN1), !(IN50 | IN47)), IN33)), IN16), (!(xor(xor(IN41 | IN9, xor(xor(IN10, false), IN32)), IN18))) & ((xor(xor(IN30 & IN49, IN35), IN49 & IN33)) & ((!(IN29)) & (xor(xor(IN45, IN43), IN26)))))), ((((IN37 | IN4) | (xor(xor(IN5, IN44), IN33))) | (xor(xor(IN40 & IN9, IN43 | IN4), xor(xor(IN41, IN16), IN9)))) | (!(IN16 | IN36))) & (!((xor(xor(IN40 | IN41, !(IN8)), xor(xor(IN50, IN30), IN14))) | (xor(xor(IN19, IN7 & IN10), xor(xor(IN24, IN40), IN28)))))))) & (xor(xor(IN22 | IN44, xor(xor(xor(xor((((!(IN12)) | IN43) | (!(!(IN46)))) & ((xor(xor(xor(xor(IN8, IN25), IN44), IN20), xor(xor(IN47, IN42), IN6))) | (xor(xor(IN1 | IN8, xor(xor(IN39, IN36), IN4)), IN11 | IN4))), (((IN28 | IN43) & (IN47 | IN33)) & IN25) & (!(IN8))), xor(xor(((IN48 & IN49) & IN49) | ((xor(xor(IN42, IN46), IN2)) | (xor(xor(IN17, IN23), IN49))), !(!(IN42))), !(!(IN43 | true)))), xor(xor(((xor(xor(IN32 | IN33, xor(xor(IN10, IN47), IN6)), !(IN32))) & IN43) | (xor(xor(!(IN3), IN4 | (xor(xor(IN30, IN34), IN17))), (IN9 | IN26) & (!(IN15)))), !(!(!(IN10 | IN23)))), xor(xor((xor(xor(IN50 | IN45, xor(xor(IN29, IN42), IN35)), IN2 & IN36)) | IN7, (IN25 & (IN24 | IN6)) & (xor(xor(IN35 & IN41, true & IN36), IN44 | IN2))), xor(xor(!(true | IN35), xor(xor(IN44 | IN41, xor(xor(IN45, IN12), IN34)), !(IN16))), !(IN2))))), !(!(!(xor(xor(IN36 & IN50, IN50), IN24 & IN9)))))), (true & (((!(IN33 | IN50)) & (!(IN2 & IN44))) | (xor(xor(IN18 & IN17, (IN21 | IN47) & (IN27 | IN27)), (IN3 & IN22) | IN49)))) & (!(xor(xor(((xor(xor(IN4, IN50), IN15)) & (IN17 | IN19)) | (!(xor(xor(IN38, IN4), IN44))), (!(!(IN16))) & IN26), ((IN20 & IN7) | (IN12 & IN31)) | (!(IN24 & IN32)))))))), (!(xor(xor(IN35, xor(xor(IN19, xor(xor(!((xor(xor(IN30, IN10), IN4)) & (IN26 & IN43)), xor(xor(xor(xor(IN8 | IN25, !(IN4)), IN26 | IN39), xor(xor(IN14, IN48 & IN29), !(IN29))), (IN47 | IN42) & IN50)), (xor(xor(true, !(IN19)), !(IN24))) & (!(IN26 & IN10)))), (IN1 & (!(xor(xor(IN2, IN27), IN47)))) & (!((IN41 & IN13) & (IN24 | IN35))))), !(IN20)))) | (!(((((!(IN36)) | IN3) | IN45) & ((((!(IN12)) | (IN49 & IN17)) | (xor(xor(!(IN49), xor(xor(IN40, IN47), IN48)), !(IN37)))) | IN40)) & (!(IN9 | (true | (!(IN44 | IN40))))))))), xor(xor(xor(xor((((!((xor(xor(!(IN15), IN45 | IN9), IN5)) & (!(IN17)))) | IN19) & (xor(xor(xor(xor(xor(xor(xor(xor(IN1, xor(xor(IN45, IN17), IN13)), xor(xor(IN9, IN3), IN47)), (IN34 | IN6) & (!(IN34))), IN6), xor(xor((!(IN41)) & (xor(xor(IN47, IN5), IN29)), !(true & IN18)), IN11)), IN49), xor(xor(IN20 | ((xor(xor(IN38, IN42), IN1)) & (!(IN39))), !((xor(xor(IN36, IN28), IN6)) | (!(IN9)))), (xor(xor(IN30, IN37 | IN9), IN12 | IN38)) | IN20)), xor(xor((IN40 | (!(IN40))) & (xor(xor(IN35 & IN45, IN15), IN18 & IN10)), !(xor(xor(xor(xor(IN11, IN42), IN31), IN2 | IN34), IN45))), (xor(xor(IN3 | IN12, IN8), IN28 | IN25)) & IN9)))) & ((IN50 | (xor(xor(!((!(IN2)) & IN29), IN4), xor(xor((xor(xor(IN33, IN15), IN27)) | (!(IN35)), xor(xor(IN11 | IN18, IN2 | true), IN19 & IN29)), (IN15 | IN6) & (IN36 | IN47))))) & IN1), xor(xor((!((((IN34 | IN23) & IN33) | ((IN26 | IN9) | (IN17 & IN17))) & (xor(xor(!(IN13 | IN4), !(IN32 | IN30)), !(IN26))))) | (((xor(xor((!(IN14)) & (!(IN28)), IN1), IN5)) | (xor(xor(xor(xor(IN24 | IN12, IN13 | false), IN21 & IN24), (IN14 | IN10) & (IN25 & IN33)), IN24))) | (IN16 & IN29)), (!(!(xor(xor(!(IN43 & IN19), !(IN26 | IN15)), (IN31 & IN23) | (xor(xor(IN28, IN20), IN7)))))) & IN17), xor(xor(((xor(xor((!(IN27)) & (IN24 & IN35), (IN40 & IN30) | (IN34 & true)), IN19)) | (IN45 | ((xor(xor(IN15, IN9), IN4)) & IN37))) | IN40, !((IN6 & (xor(xor(xor(xor(IN3, IN9), IN33), !(IN47)), IN39 & IN5))) & (xor(xor(IN36, xor(xor(false | IN47, xor(xor(IN24, IN35), IN1)), IN45 & IN13)), (!(IN36)) | (IN38 & IN3))))), (xor(xor(IN35, (!(!(IN43))) | ((!(IN4)) | (xor(xor(IN9, IN19), IN36)))), xor(xor(IN38, xor(xor(xor(xor(IN48, IN41), IN7), IN30), !(IN24))), !(!(IN8))))) & (xor(xor(((IN34 | IN24) & (!(IN44))) | (!(IN42 | IN34)), xor(xor(xor(xor(IN16 & IN19, IN33), xor(xor(IN5, IN3), IN19)), IN34), IN19 | (IN3 | IN7))), xor(xor(IN43, xor(xor(false | IN25, IN16 & IN14), IN31 & IN6)), xor(xor(IN5, xor(xor(IN35, IN17), IN2)), IN8 & IN22))))))), IN9), IN41 | (!(!(xor(xor((!(!(!(IN36)))) | (!(!(xor(xor(IN4, IN32), IN32)))), xor(xor(IN13, (xor(xor(IN19, IN38 & IN33), !(IN41))) | (!(!(IN39)))), IN9)), xor(xor(IN29, !((true & IN12) | (xor(xor(IN3, false), IN35)))), ((xor(xor(IN10, IN19), IN7)) | (IN2 | true)) | IN48)))))), ((xor(xor(!(xor(xor(!((IN35 | IN36) & (IN15 & IN44)), xor(xor((xor(xor(IN37, IN25), IN10)) & IN12, !(!(IN46))), !(IN37 | IN9))), ((IN2 & IN19) & (IN1 | IN6)) | (!(IN1 & IN20)))), xor(xor((!(!(IN1 & IN39))) & IN32, xor(xor(!(xor(xor(IN9 | IN11, IN13 & IN43), !(IN29))), xor(xor(IN50 | true, !(IN36 & IN13)), (!(IN20)) | IN50)), xor(xor(IN12 | (xor(xor(IN19, IN15), IN32)), xor(xor(IN34 | IN5, !(IN19)), IN33 | IN43)), xor(xor(IN18 & IN17, IN22), xor(xor(IN41, IN30), IN28))))), !((!(!(IN47))) | (!(IN14))))), xor(xor(IN5, IN10), (!(IN13)) | IN35))) & IN11) & (xor(xor((!((!((!(IN35)) & IN47)) & IN28)) | (xor(xor((IN16 & (IN24 & (IN49 & IN16))) & IN41, ((!(xor(xor(IN18, IN33), IN30))) | ((IN13 & IN44) | (xor(xor(IN21, IN38), IN2)))) | ((!(IN38)) | (!(IN25 & IN24)))), xor(xor(!((!(IN13)) | IN5), (!(IN24)) & ((IN44 | IN13) | (xor(xor(IN13, IN6), IN19)))), xor(xor((IN36 & IN49) | true, !(IN4 & IN35)), xor(xor(IN25 & IN13, IN41), xor(xor(IN16, IN26), false)))))), IN27), !(IN42)))))

*)

FUNCTION_BLOCK F_CollectInput
  VAR_IN_OUT
      Data : ARRAY[1..50] OF BOOL;
  END_VAR
  VAR_INPUT
      TICK  : BOOL := 0;
      IN1   : BOOL := 0;
      IN2   : BOOL := 0;
      IN3   : BOOL := 0;
      IN4   : BOOL := 0;
      IN5   : BOOL := 0;
      RESET : BOOL := FALSE;
  END_VAR
  VAR_OUTPUT
      Finished : BOOL;
  END_VAR
  VAR
      j    : USINT := 1;
      tock : BOOL  := 0;
  END_VAR
  IF NOT RESET AND tock = NOT TICK THEN
      Data[j]   := IN1;
      Data[j+1] := IN2;
      Data[j+2] := IN3;
      Data[j+3] := IN4;
      Data[j+4] := IN5;
      j := j + 5;
      tock := TICK;
  ELSE
      j := 1;
      tock := 0;
  END_IF;
  Finished := (j > 50);
END_FUNCTION_BLOCK

PROGRAM Boiler
  VAR
    Data  : ARRAY[1..50] OF BOOL;
    Ready : BOOL;
    CollectInput : F_CollectInput;
  END_VAR
  VAR
    TICK     AT %IX1.0 : BOOL;
    IN1      AT %IX0.3 : BOOL;
    IN2      AT %IX0.4 : BOOL;
    IN3      AT %IX0.5 : BOOL;
    IN4      AT %IX0.6 : BOOL;
    IN5      AT %IX0.7 : BOOL;
    OutReady AT %QX0.0 : BOOL := FALSE;
    FeedNext AT %QX0.1 : BOOL := FALSE;
    Out      AT %QX0.2 : BOOL;
  END_VAR
  CollectInput(TICK:=TICK, IN1:=IN1, IN2:=IN2, IN3:=IN3, IN4:=IN4, IN5:=IN5);
  Ready := CollectInput.Finished;
  FeedNext := 1;
  IF Ready THEN
    Out := ((((Data[21] XOR ((Data[18] AND ((((((((Data[50] OR Data[1]) AND (Data[14] AND Data[11])) XOR (((Data[43] OR Data[14]) XOR ((Data[44] XOR Data[33]) XOR Data[13])) XOR (NOT Data[12]))) XOR Data[23]) OR ((((NOT Data[4]) AND (NOT Data[36])) XOR ((Data[18] OR Data[26]) OR (Data[35] OR Data[4]))) XOR Data[17])) OR (Data[48] OR (NOT (((Data[18] XOR Data[37]) XOR Data[11]) OR Data[15])))) XOR (Data[14] AND (NOT Data[48]))) XOR (Data[43] AND ((((((NOT Data[37]) AND (Data[28] AND Data[40])) XOR Data[2]) XOR ((NOT Data[3]) OR (Data[40] AND Data[12]))) XOR (((((Data[28] AND Data[23]) XOR Data[41]) XOR (NOT Data[32])) XOR ((NOT Data[47]) AND (NOT Data[32]))) XOR ((NOT Data[12]) OR ((Data[29] XOR FALSE) XOR Data[29])))) XOR (((((NOT Data[14]) XOR (NOT Data[13])) XOR (Data[21] OR Data[22])) XOR (((NOT Data[43]) XOR (Data[19] OR Data[33])) XOR ((Data[36] XOR Data[14]) XOR Data[24]))) XOR TRUE))))) AND ((Data[35] OR Data[16]) OR Data[50]))) XOR ((Data[42] XOR Data[33]) XOR Data[47])) XOR (((((NOT (((((Data[10] OR ((Data[36] XOR Data[36]) XOR Data[48])) OR ((NOT Data[42]) AND (Data[8] OR Data[31]))) XOR (((NOT Data[11]) OR (Data[12] AND Data[9])) OR (((Data[8] XOR Data[5]) XOR Data[3]) OR (TRUE OR Data[26])))) XOR (NOT ((Data[24] OR Data[50]) AND ((Data[15] XOR Data[45]) XOR Data[38])))) AND (((Data[42] OR ((Data[18] OR Data[37]) AND (Data[15] AND Data[43]))) XOR ((NOT Data[15]) OR ((Data[25] OR Data[45]) OR ((Data[19] XOR Data[35]) XOR Data[4])))) XOR (Data[3] OR (NOT (Data[13] OR Data[38])))))) OR (Data[14] OR ((((((NOT Data[1]) OR (Data[2] AND Data[27])) AND ((Data[45] OR Data[39]) AND FALSE)) XOR (((NOT (NOT Data[21])) XOR Data[27]) XOR ((Data[19] OR Data[19]) OR (Data[14] OR Data[32])))) XOR (((((TRUE XOR Data[5]) XOR Data[21]) XOR ((Data[38] XOR Data[6]) XOR Data[18])) XOR ((Data[2] XOR Data[3]) XOR TRUE)) AND (NOT (Data[44] AND Data[27])))) OR (NOT (((Data[5] AND Data[37]) AND Data[1]) OR ((Data[18] AND Data[28]) AND (Data[33] OR Data[49]))))))) OR (NOT (NOT ((NOT Data[26]) OR (NOT ((((Data[23] OR Data[42]) XOR (NOT Data[8])) XOR (NOT Data[5])) AND ((Data[8] AND Data[13]) AND ((Data[36] XOR Data[2]) XOR Data[28])))))))) XOR (((Data[48] XOR (((Data[37] AND ((Data[8] XOR Data[38]) XOR ((NOT (Data[20] OR Data[8])) OR ((Data[32] OR Data[43]) AND (NOT Data[9]))))) XOR ((NOT (Data[28] OR (((Data[40] AND Data[12]) XOR (NOT Data[46])) XOR (Data[17] AND Data[49])))) OR Data[38])) XOR Data[3])) XOR (((NOT (NOT (((((NOT Data[23]) XOR Data[1]) XOR (Data[18] AND Data[50])) XOR (NOT (NOT Data[11]))) XOR ((((Data[47] XOR Data[15]) XOR Data[49]) XOR (NOT Data[44])) XOR (NOT Data[44]))))) XOR ((((((NOT (Data[29] OR Data[44])) OR Data[43]) XOR Data[34]) XOR (((((Data[8] AND Data[46]) XOR Data[14]) XOR (Data[25] AND Data[1])) XOR (NOT (Data[50] OR Data[47]))) XOR Data[33])) XOR Data[16]) XOR ((NOT (((Data[41] OR Data[9]) XOR ((Data[10] XOR FALSE) XOR Data[32])) XOR Data[18])) AND ((((Data[30] AND Data[49]) XOR Data[35]) XOR (Data[49] AND Data[33])) AND ((NOT Data[29]) AND ((Data[45] XOR Data[43]) XOR Data[26])))))) XOR (((((Data[37] OR Data[4]) OR ((Data[5] XOR Data[44]) XOR Data[33])) OR (((Data[40] AND Data[9]) XOR (Data[43] OR Data[4])) XOR ((Data[41] XOR Data[16]) XOR Data[9]))) OR (NOT (Data[16] OR Data[36]))) AND (NOT ((((Data[40] OR Data[41]) XOR (NOT Data[8])) XOR ((Data[50] XOR Data[30]) XOR Data[14])) OR ((Data[19] XOR (Data[7] AND Data[10])) XOR ((Data[24] XOR Data[40]) XOR Data[28]))))))) AND (((Data[22] OR Data[44]) XOR ((((((((NOT Data[12]) OR Data[43]) OR (NOT (NOT Data[46]))) AND (((((Data[8] XOR Data[25]) XOR Data[44]) XOR Data[20]) XOR ((Data[47] XOR Data[42]) XOR Data[6])) OR (((Data[1] OR Data[8]) XOR ((Data[39] XOR Data[36]) XOR Data[4])) XOR (Data[11] OR Data[4])))) XOR ((((Data[28] OR Data[43]) AND (Data[47] OR Data[33])) AND Data[25]) AND (NOT Data[8]))) XOR (((((Data[48] AND Data[49]) AND Data[49]) OR (((Data[42] XOR Data[46]) XOR Data[2]) OR ((Data[17] XOR Data[23]) XOR Data[49]))) XOR (NOT (NOT Data[42]))) XOR (NOT (NOT (Data[43] OR TRUE))))) XOR (((((((Data[32] OR Data[33]) XOR ((Data[10] XOR Data[47]) XOR Data[6])) XOR (NOT Data[32])) AND Data[43]) OR (((NOT Data[3]) XOR (Data[4] OR ((Data[30] XOR Data[34]) XOR Data[17]))) XOR ((Data[9] OR Data[26]) AND (NOT Data[15])))) XOR (NOT (NOT (NOT (Data[10] OR Data[23]))))) XOR ((((((Data[50] OR Data[45]) XOR ((Data[29] XOR Data[42]) XOR Data[35])) XOR (Data[2] AND Data[36])) OR Data[7]) XOR ((Data[25] AND (Data[24] OR Data[6])) AND (((Data[35] AND Data[41]) XOR (TRUE AND Data[36])) XOR (Data[44] OR Data[2])))) XOR (((NOT (TRUE OR Data[35])) XOR (((Data[44] OR Data[41]) XOR ((Data[45] XOR Data[12]) XOR Data[34])) XOR (NOT Data[16]))) XOR (NOT Data[2]))))) XOR (NOT (NOT (NOT (((Data[36] AND Data[50]) XOR Data[50]) XOR (Data[24] AND Data[9]))))))) XOR ((TRUE AND (((NOT (Data[33] OR Data[50])) AND (NOT (Data[2] AND Data[44]))) OR (((Data[18] AND Data[17]) XOR ((Data[21] OR Data[47]) AND (Data[27] OR Data[27]))) XOR ((Data[3] AND Data[22]) OR Data[49])))) AND (NOT ((((((Data[4] XOR Data[50]) XOR Data[15]) AND (Data[17] OR Data[19])) OR (NOT ((Data[38] XOR Data[4]) XOR Data[44]))) XOR ((NOT (NOT Data[16])) AND Data[26])) XOR (((Data[20] AND Data[7]) OR (Data[12] AND Data[31])) OR (NOT (Data[24] AND Data[32]))))))))) XOR ((NOT ((Data[35] XOR ((Data[19] XOR (((NOT (((Data[30] XOR Data[10]) XOR Data[4]) AND (Data[26] AND Data[43]))) XOR (((((Data[8] OR Data[25]) XOR (NOT Data[4])) XOR (Data[26] OR Data[39])) XOR ((Data[14] XOR (Data[48] AND Data[29])) XOR (NOT Data[29]))) XOR ((Data[47] OR Data[42]) AND Data[50]))) XOR (((TRUE XOR (NOT Data[19])) XOR (NOT Data[24])) AND (NOT (Data[26] AND Data[10]))))) XOR ((Data[1] AND (NOT ((Data[2] XOR Data[27]) XOR Data[47]))) AND (NOT ((Data[41] AND Data[13]) AND (Data[24] OR Data[35])))))) XOR (NOT Data[20]))) OR (NOT (((((NOT Data[36]) OR Data[3]) OR Data[45]) AND ((((NOT Data[12]) OR (Data[49] AND Data[17])) OR (((NOT Data[49]) XOR ((Data[40] XOR Data[47]) XOR Data[48])) XOR (NOT Data[37]))) OR Data[40])) AND (NOT (Data[9] OR (TRUE OR (NOT (Data[44] OR Data[40])))))))))) XOR ((((((((NOT ((((NOT Data[15]) XOR (Data[45] OR Data[9])) XOR Data[5]) AND (NOT Data[17]))) OR Data[19]) AND ((((((((Data[1] XOR ((Data[45] XOR Data[17]) XOR Data[13])) XOR ((Data[9] XOR Data[3]) XOR Data[47])) XOR ((Data[34] OR Data[6]) AND (NOT Data[34]))) XOR Data[6]) XOR ((((NOT Data[41]) AND ((Data[47] XOR Data[5]) XOR Data[29])) XOR (NOT (TRUE AND Data[18]))) XOR Data[11])) XOR Data[49]) XOR (((Data[20] OR (((Data[38] XOR Data[42]) XOR Data[1]) AND (NOT Data[39]))) XOR (NOT (((Data[36] XOR Data[28]) XOR Data[6]) OR (NOT Data[9])))) XOR (((Data[30] XOR (Data[37] OR Data[9])) XOR (Data[12] OR Data[38])) OR Data[20]))) XOR ((((Data[40] OR (NOT Data[40])) AND (((Data[35] AND Data[45]) XOR Data[15]) XOR (Data[18] AND Data[10]))) XOR (NOT ((((Data[11] XOR Data[42]) XOR Data[31]) XOR (Data[2] OR Data[34])) XOR Data[45]))) XOR ((((Data[3] OR Data[12]) XOR Data[8]) XOR (Data[28] OR Data[25])) AND Data[9])))) AND ((Data[50] OR (((NOT ((NOT Data[2]) AND Data[29])) XOR Data[4]) XOR (((((Data[33] XOR Data[15]) XOR Data[27]) OR (NOT Data[35])) XOR (((Data[11] OR Data[18]) XOR (Data[2] OR TRUE)) XOR (Data[19] AND Data[29]))) XOR ((Data[15] OR Data[6]) AND (Data[36] OR Data[47]))))) AND Data[1])) XOR ((((NOT ((((Data[34] OR Data[23]) AND Data[33]) OR ((Data[26] OR Data[9]) OR (Data[17] AND Data[17]))) AND (((NOT (Data[13] OR Data[4])) XOR (NOT (Data[32] OR Data[30]))) XOR (NOT Data[26])))) OR ((((((NOT Data[14]) AND (NOT Data[28])) XOR Data[1]) XOR Data[5]) OR (((((Data[24] OR Data[12]) XOR (Data[13] OR FALSE)) XOR (Data[21] AND Data[24])) XOR ((Data[14] OR Data[10]) AND (Data[25] AND Data[33]))) XOR Data[24])) OR (Data[16] AND Data[29]))) XOR ((NOT (NOT (((NOT (Data[43] AND Data[19])) XOR (NOT (Data[26] OR Data[15]))) XOR ((Data[31] AND Data[23]) OR ((Data[28] XOR Data[20]) XOR Data[7]))))) AND Data[17])) XOR ((((((((NOT Data[27]) AND (Data[24] AND Data[35])) XOR ((Data[40] AND Data[30]) OR (Data[34] AND TRUE))) XOR Data[19]) OR (Data[45] OR (((Data[15] XOR Data[9]) XOR Data[4]) AND Data[37]))) OR Data[40]) XOR (NOT ((Data[6] AND ((((Data[3] XOR Data[9]) XOR Data[33]) XOR (NOT Data[47])) XOR (Data[39] AND Data[5]))) AND ((Data[36] XOR (((FALSE OR Data[47]) XOR ((Data[24] XOR Data[35]) XOR Data[1])) XOR (Data[45] AND Data[13]))) XOR ((NOT Data[36]) OR (Data[38] AND Data[3])))))) XOR (((Data[35] XOR ((NOT (NOT Data[43])) OR ((NOT Data[4]) OR ((Data[9] XOR Data[19]) XOR Data[36])))) XOR ((Data[38] XOR ((((Data[48] XOR Data[41]) XOR Data[7]) XOR Data[30]) XOR (NOT Data[24]))) XOR (NOT (NOT Data[8])))) AND (((((Data[34] OR Data[24]) AND (NOT Data[44])) OR (NOT (Data[42] OR Data[34]))) XOR (((((Data[16] AND Data[19]) XOR Data[33]) XOR ((Data[5] XOR Data[3]) XOR Data[19])) XOR Data[34]) XOR (Data[19] OR (Data[3] OR Data[7])))) XOR ((Data[43] XOR (((FALSE OR Data[25]) XOR (Data[16] AND Data[14])) XOR (Data[31] AND Data[6]))) XOR ((Data[5] XOR ((Data[35] XOR Data[17]) XOR Data[2])) XOR (Data[8] AND Data[22])))))))) XOR Data[9]) XOR (Data[41] OR (NOT (NOT ((((NOT (NOT (NOT Data[36]))) OR (NOT (NOT ((Data[4] XOR Data[32]) XOR Data[32])))) XOR ((Data[13] XOR (((Data[19] XOR (Data[38] AND Data[33])) XOR (NOT Data[41])) OR (NOT (NOT Data[39])))) XOR Data[9])) XOR ((Data[29] XOR (NOT ((TRUE AND Data[12]) OR ((Data[3] XOR FALSE) XOR Data[35])))) XOR ((((Data[10] XOR Data[19]) XOR Data[7]) OR (Data[2] OR TRUE)) OR Data[48]))))))) XOR (((((NOT (((NOT ((Data[35] OR Data[36]) AND (Data[15] AND Data[44]))) XOR (((((Data[37] XOR Data[25]) XOR Data[10]) AND Data[12]) XOR (NOT (NOT Data[46]))) XOR (NOT (Data[37] OR Data[9])))) XOR (((Data[2] AND Data[19]) AND (Data[1] OR Data[6])) OR (NOT (Data[1] AND Data[20]))))) XOR ((((NOT (NOT (Data[1] AND Data[39]))) AND Data[32]) XOR (((NOT (((Data[9] OR Data[11]) XOR (Data[13] AND Data[43])) XOR (NOT Data[29]))) XOR (((Data[50] OR TRUE) XOR (NOT (Data[36] AND Data[13]))) XOR ((NOT Data[20]) OR Data[50]))) XOR (((Data[12] OR ((Data[19] XOR Data[15]) XOR Data[32])) XOR (((Data[34] OR Data[5]) XOR (NOT Data[19])) XOR (Data[33] OR Data[43]))) XOR (((Data[18] AND Data[17]) XOR Data[22]) XOR ((Data[41] XOR Data[30]) XOR Data[28]))))) XOR (NOT ((NOT (NOT Data[47])) OR (NOT Data[14]))))) XOR ((Data[5] XOR Data[10]) XOR ((NOT Data[13]) OR Data[35]))) AND Data[11]) AND ((((NOT ((NOT ((NOT Data[35]) AND Data[47])) AND Data[28])) OR ((((Data[16] AND (Data[24] AND (Data[49] AND Data[16]))) AND Data[41]) XOR (((NOT ((Data[18] XOR Data[33]) XOR Data[30])) OR ((Data[13] AND Data[44]) OR ((Data[21] XOR Data[38]) XOR Data[2]))) OR ((NOT Data[38]) OR (NOT (Data[25] AND Data[24]))))) XOR (((NOT ((NOT Data[13]) OR Data[5])) XOR ((NOT Data[24]) AND ((Data[44] OR Data[13]) OR ((Data[13] XOR Data[6]) XOR Data[19])))) XOR ((((Data[36] AND Data[49]) OR TRUE) XOR (NOT (Data[4] AND Data[35]))) XOR (((Data[25] AND Data[13]) XOR Data[41]) XOR ((Data[16] XOR Data[26]) XOR FALSE)))))) XOR Data[27]) XOR (NOT Data[42])))));
    OutReady := 1;
    CollectInput(RESET:=TRUE);
  END_IF;
END_PROGRAM

CONFIGURATION Config0
  RESOURCE Res0 ON PLC
    TASK task0(INTERVAL := T#20ms,PRIORITY := 0);
    PROGRAM instance0 WITH task0 : Boiler;
  END_RESOURCE
END_CONFIGURATION

(* ---- RND-EXPR_linty-mujik-lodge.st ---- *)
(*
This code implements a randomly grown symbolic expression:

xor(xor(xor(xor(xor(xor((xor(xor(xor(xor(IN26, !(IN6)), (((IN11 | IN7) | (IN46 | IN35)) & ((xor(xor(IN35, IN31), IN1)) | (IN42 & IN18))) & (((IN36 & IN18) | (xor(xor(IN36, IN17), IN50))) & (!(IN12 & IN48)))), xor(xor((xor(xor(xor(xor(IN10 | IN24, IN32 | IN19), !(IN47)), (IN10 & IN32) | (IN28 | IN34)), !(xor(xor(IN29, IN40), IN46)))) | (((xor(xor(IN29, IN25), IN6)) | (IN31 | IN35)) & (xor(xor(!(IN7), xor(xor(IN38, IN3), IN32)), IN36))), IN35), xor(xor((xor(xor(IN1 & IN29, !(IN2)), IN21 & IN10)) | IN34, IN22 | IN29), xor(xor((!(IN25)) & (!(IN13)), (IN20 | IN2) | (!(IN4))), IN10)))), (((!(xor(xor(IN41, IN6), IN14))) | ((xor(xor(IN9, IN5), IN35)) & (xor(xor(true, IN31), IN11)))) & ((xor(xor(IN35 | IN15, IN32 | IN26), IN12 | IN43)) | IN4)) | ((xor(xor((IN44 | IN44) & (xor(xor(IN28, IN43), IN17)), IN44), !(IN9 & IN28))) & (xor(xor(IN29 | (IN30 | IN27), xor(xor(IN27, xor(xor(true, IN9), IN43)), IN6 | IN39)), IN46 | (!(IN39))))))) | ((!(IN9)) | (!(xor(xor(IN42, IN9 | (xor(xor(IN38 & IN48, xor(xor(IN22, IN35), IN3)), xor(xor(IN19, IN27), IN18)))), IN1)))), ((!(IN47)) & ((!(xor(xor(!(IN5), xor(xor(!(IN12), IN14), xor(xor(IN25, IN40), IN25))), !(xor(xor(false, IN36), IN17))))) | (!(xor(xor(xor(xor(xor(xor(IN25, IN10), IN29), IN38 & IN2), !(IN29)), (IN41 | IN2) | (IN16 | IN26)), (xor(xor(IN44, IN2), IN33)) & (IN25 & IN25)))))) | (xor(xor(xor(xor(IN35 & (xor(xor((xor(xor(IN46, IN22), IN20)) & (IN19 | IN9), IN45), !(IN40 | IN20))), !(!(!(IN16 | IN30)))), xor(xor(IN29 & (xor(xor(xor(xor(IN34, IN31), IN16), xor(xor(IN24, IN10), IN20)), !(IN8))), ((IN30 | IN45) | IN15) | (xor(xor(!(IN38), IN46 | IN14), !(IN2)))), IN25)), xor(xor(IN26, !(IN39 | ((!(IN11)) & (!(IN12))))), IN31)), (((xor(xor(xor(xor(IN44, IN49), IN41), IN22 | IN11), xor(xor(IN1, IN15), IN32))) & (IN43 & (IN50 & IN31))) & (((!(IN7)) & (xor(xor(IN46, IN41), IN40))) | (!(IN12 | IN11)))) & (!(((IN34 & IN11) & (IN42 | IN24)) & ((IN21 | IN4) | (xor(xor(IN23, IN28), IN40)))))))), xor(xor((((((!(IN20)) & (IN30 | IN35)) & (xor(xor(xor(xor(true, IN30), IN21), IN30 & IN39), IN20 | IN26))) | (IN48 & ((!(IN37)) | IN31))) | ((((!(IN26)) & (IN20 & IN29)) & ((!(IN28)) | IN14)) & (IN32 & ((IN34 | IN42) & (IN47 & IN46))))) & (!(IN41)), IN50), IN28 | (!(false | (xor(xor(xor(xor(IN16 | true, IN48 | IN47), xor(xor(IN45, IN16), IN31)), xor(xor(xor(xor(false, IN18), IN37), IN46), IN28 | IN12)), (IN45 & IN4) & (!(IN31)))))))), xor(xor(!(((!(!(IN19))) | ((IN30 | (!(xor(xor(IN36, IN3), IN50)))) & IN31)) & IN8), ((!(!(((IN35 & IN23) | (IN40 | IN11)) | ((xor(xor(IN12, IN42), IN32)) | (!(IN34)))))) & (!(IN7))) & ((IN15 & IN27) & ((xor(xor(!(xor(xor(!(IN12), !(IN21)), IN39 | IN21)), (!(xor(xor(IN31, IN26), IN50))) | (xor(xor(xor(xor(IN7, IN6), IN11), IN18), IN4))), xor(xor((!(IN28)) & (xor(xor(IN19, IN4), IN16)), xor(xor(!(IN23), xor(xor(IN34, IN42), IN15)), xor(xor(IN40, IN20), true))), (!(IN6)) | (IN12 & IN2)))) | (!(xor(xor(IN46, (IN14 & IN43) & IN50), IN6)))))), (!(!((xor(xor(IN49, (IN10 & IN41) & (false & IN10)), xor(xor(xor(xor(IN38, IN33), IN36), IN29 & IN4), IN43))) & (!((!(IN3)) & IN9))))) & (!(IN5)))), ((!((!(((!(IN6)) & (IN1 | IN28)) & (!(xor(xor(IN26, IN28), IN16))))) & (xor(xor(!(IN18), IN22), ((IN20 & IN15) | (!(IN40))) & (!(IN2 & IN7)))))) | ((xor(xor((((IN50 | IN5) & IN50) & (xor(xor(!(IN40), IN18 | IN38), !(IN31)))) | IN48, xor(xor((xor(xor(xor(xor(IN15, IN26), IN23), IN33 | IN44), IN6)) & (!(xor(xor(IN35, IN26), IN47))), ((!(IN7)) & (!(IN14))) & (IN33 | IN50)), IN48)), !(IN32 | (!(IN20 | IN48))))) & (xor(xor(((IN16 | (!(IN1))) | (!(IN46 & IN16))) & (((!(IN2)) | (IN36 & IN9)) | ((IN4 & IN34) & (IN37 | IN13))), IN23), IN4 | (IN27 | (xor(xor(IN35 | IN31, IN9 | IN11), IN23 & IN37))))))) & (((IN22 | (((xor(xor(!(IN32), xor(xor(IN24, IN27), IN47)), IN32)) | ((!(IN37)) | (!(IN46)))) & IN28)) & (!(IN8 | (((!(IN42)) | (IN46 | IN24)) & ((!(IN33)) & (xor(xor(IN25, IN24), IN9))))))) | (((((IN26 & IN8) & IN49) | (!(IN2))) & (((xor(xor(IN7, xor(xor(IN25, IN31), IN21)), !(IN38))) | ((IN29 | IN14) & (IN34 | IN25))) & ((!(xor(xor(IN18, IN6), IN48))) & IN7))) | IN13))), IN37), ((!(xor(xor(IN15, !((((!(IN46)) | (IN25 | IN41)) | (xor(xor(false | IN14, xor(xor(IN27, IN2), IN33)), !(IN33)))) & IN17)), IN37 | (xor(xor(!((IN24 | IN45) | (xor(xor(IN33, IN46), IN36))), ((!(IN10)) | (IN10 | IN28)) | ((IN3 | IN26) & IN48)), ((IN14 & true) & (!(IN17))) | ((!(IN50)) | (IN48 & true))))))) & IN17) | (xor(xor(!((xor(xor(xor(xor(IN30 | ((IN12 | IN23) & IN24), (xor(xor(IN13, IN11), IN1)) | (!(IN38))), IN39 & (!(xor(xor(IN3, IN20), IN5)))), IN21 | ((!(IN33 | IN7)) | IN31)), !(!(IN49)))) | IN41), xor(xor(true, xor(xor((xor(xor(IN39, xor(xor((IN17 & IN5) & IN4, !(IN49 & IN25)), !(IN39))), IN32)) | (!(IN6 & IN44)), (((IN18 | (!(IN31))) & ((!(IN48)) | (IN21 | IN41))) | IN20) & ((!((!(IN28)) & (xor(xor(IN18, IN44), IN40)))) | (IN12 | (xor(xor(IN5 | IN13, IN48 | IN34), IN30))))), IN23)), IN45)), ((xor(xor(!(!(IN44)), (xor(xor((xor(xor(false, IN24), IN5)) | (xor(xor(IN27, IN9), IN19)), xor(xor(IN47, xor(xor(IN17, IN1), IN11)), IN34)), !(xor(xor(IN23, IN47), IN23)))) & (xor(xor(IN7 | (xor(xor(IN36, true), IN6)), (xor(xor(IN5, IN2), IN29)) | (xor(xor(IN1, IN46), IN47))), (IN40 & IN29) & (xor(xor(IN38, IN44), false))))), ((xor(xor(IN2 | IN12, IN1 | IN17), xor(xor(IN17, IN4), IN32))) | ((xor(xor(IN19, IN41), IN36)) | (IN18 | IN5))) | IN16)) | (IN45 | (!(xor(xor(IN26, !(IN22 & IN9)), (IN28 | IN40) | (xor(xor(IN39, IN15), IN21))))))) & (!(IN24 | ((((IN38 | IN48) | (IN8 & IN6)) & (xor(xor(xor(xor(IN38, IN9), IN11), IN44 & IN3), IN11 | IN50))) | (((!(IN30)) & (IN37 & IN27)) | ((!(IN5)) & (IN34 & IN22)))))))))

*)

FUNCTION_BLOCK F_CollectInput
  VAR_IN_OUT
      Data : ARRAY[1..50] OF BOOL;
  END_VAR
  VAR_INPUT
      TICK  : BOOL := 0;
      IN1   : BOOL := 0;
      IN2   : BOOL := 0;
      IN3   : BOOL := 0;
      IN4   : BOOL := 0;
      IN5   : BOOL := 0;
      RESET : BOOL := FALSE;
  END_VAR
  VAR_OUTPUT
      Finished : BOOL;
  END_VAR
  VAR
      j    : USINT := 1;
      tock : BOOL  := 0;
  END_VAR
  IF NOT RESET AND tock = NOT TICK THEN
      Data[j]   := IN1;
      Data[j+1] := IN2;
      Data[j+2] := IN3;
      Data[j+3] := IN4;
      Data[j+4] := IN5;
      j := j + 5;
      tock := TICK;
  ELSE
      j := 1;
      tock := 0;
  END_IF;
  Finished := (j > 50);
END_FUNCTION_BLOCK

PROGRAM Boiler
  VAR
    Data  : ARRAY[1..50] OF BOOL;
    Ready : BOOL;
    CollectInput : F_CollectInput;
  END_VAR
  VAR
    TICK     AT %IX1.0 : BOOL;
    IN1      AT %IX0.3 : BOOL;
    IN2      AT %IX0.4 : BOOL;
    IN3      AT %IX0.5 : BOOL;
    IN4      AT %IX0.6 : BOOL;
    IN5      AT %IX0.7 : BOOL;
    OutReady AT %QX0.0 : BOOL := FALSE;
    FeedNext AT %QX0.1 : BOOL := FALSE;
    Out      AT %QX0.2 : BOOL;
  END_VAR
  CollectInput(TICK:=TICK, IN1:=IN1, IN2:=IN2, IN3:=IN3, IN4:=IN4, IN5:=IN5);
  Ready := CollectInput.Finished;
  FeedNext := 1;
  IF Ready THEN
    Out := (((((((((((Data[26] XOR (NOT Data[6])) XOR ((((Data[11] OR Data[7]) OR (Data[46] OR Data[35])) AND (((Data[35] XOR Data[31]) XOR Data[1]) OR (Data[42] AND Data[18]))) AND (((Data[36] AND Data[18]) OR ((Data[36] XOR Data[17]) XOR Data[50])) AND (NOT (Data[12] AND Data[48]))))) XOR ((((((((Data[10] OR Data[24]) XOR (Data[32] OR Data[19])) XOR (NOT Data[47])) XOR ((Data[10] AND Data[32]) OR (Data[28] OR Data[34]))) XOR (NOT ((Data[29] XOR Data[40]) XOR Data[46]))) OR ((((Data[29] XOR Data[25]) XOR Data[6]) OR (Data[31] OR Data[35])) AND (((NOT Data[7]) XOR ((Data[38] XOR Data[3]) XOR Data[32])) XOR Data[36]))) XOR Data[35]) XOR ((((((Data[1] AND Data[29]) XOR (NOT Data[2])) XOR (Data[21] AND Data[10])) OR Data[34]) XOR (Data[22] OR Data[29])) XOR ((((NOT Data[25]) AND (NOT Data[13])) XOR ((Data[20] OR Data[2]) OR (NOT Data[4]))) XOR Data[10])))) XOR ((((NOT ((Data[41] XOR Data[6]) XOR Data[14])) OR (((Data[9] XOR Data[5]) XOR Data[35]) AND ((TRUE XOR Data[31]) XOR Data[11]))) AND ((((Data[35] OR Data[15]) XOR (Data[32] OR Data[26])) XOR (Data[12] OR Data[43])) OR Data[4])) OR (((((Data[44] OR Data[44]) AND ((Data[28] XOR Data[43]) XOR Data[17])) XOR Data[44]) XOR (NOT (Data[9] AND Data[28]))) AND (((Data[29] OR (Data[30] OR Data[27])) XOR ((Data[27] XOR ((TRUE XOR Data[9]) XOR Data[43])) XOR (Data[6] OR Data[39]))) XOR (Data[46] OR (NOT Data[39])))))) OR ((NOT Data[9]) OR (NOT ((Data[42] XOR (Data[9] OR (((Data[38] AND Data[48]) XOR ((Data[22] XOR Data[35]) XOR Data[3])) XOR ((Data[19] XOR Data[27]) XOR Data[18])))) XOR Data[1])))) XOR (((NOT Data[47]) AND ((NOT (((NOT Data[5]) XOR (((NOT Data[12]) XOR Data[14]) XOR ((Data[25] XOR Data[40]) XOR Data[25]))) XOR (NOT ((FALSE XOR Data[36]) XOR Data[17])))) OR (NOT ((((((Data[25] XOR Data[10]) XOR Data[29]) XOR (Data[38] AND Data[2])) XOR (NOT Data[29])) XOR ((Data[41] OR Data[2]) OR (Data[16] OR Data[26]))) XOR (((Data[44] XOR Data[2]) XOR Data[33]) AND (Data[25] AND Data[25])))))) OR (((((Data[35] AND (((((Data[46] XOR Data[22]) XOR Data[20]) AND (Data[19] OR Data[9])) XOR Data[45]) XOR (NOT (Data[40] OR Data[20])))) XOR (NOT (NOT (NOT (Data[16] OR Data[30]))))) XOR (((Data[29] AND ((((Data[34] XOR Data[31]) XOR Data[16]) XOR ((Data[24] XOR Data[10]) XOR Data[20])) XOR (NOT Data[8]))) XOR (((Data[30] OR Data[45]) OR Data[15]) OR (((NOT Data[38]) XOR (Data[46] OR Data[14])) XOR (NOT Data[2])))) XOR Data[25])) XOR ((Data[26] XOR (NOT (Data[39] OR ((NOT Data[11]) AND (NOT Data[12]))))) XOR Data[31])) XOR (((((((Data[44] XOR Data[49]) XOR Data[41]) XOR (Data[22] OR Data[11])) XOR ((Data[1] XOR Data[15]) XOR Data[32])) AND (Data[43] AND (Data[50] AND Data[31]))) AND (((NOT Data[7]) AND ((Data[46] XOR Data[41]) XOR Data[40])) OR (NOT (Data[12] OR Data[11])))) AND (NOT (((Data[34] AND Data[11]) AND (Data[42] OR Data[24])) AND ((Data[21] OR Data[4]) OR ((Data[23] XOR Data[28]) XOR Data[40])))))))) XOR ((((((((NOT Data[20]) AND (Data[30] OR Data[35])) AND ((((TRUE XOR Data[30]) XOR Data[21]) XOR (Data[30] AND Data[39])) XOR (Data[20] OR Data[26]))) OR (Data[48] AND ((NOT Data[37]) OR Data[31]))) OR ((((NOT Data[26]) AND (Data[20] AND Data[29])) AND ((NOT Data[28]) OR Data[14])) AND (Data[32] AND ((Data[34] OR Data[42]) AND (Data[47] AND Data[46]))))) AND (NOT Data[41])) XOR Data[50]) XOR (Data[28] OR (NOT (FALSE OR (((((Data[16] OR TRUE) XOR (Data[48] OR Data[47])) XOR ((Data[45] XOR Data[16]) XOR Data[31])) XOR ((((FALSE XOR Data[18]) XOR Data[37]) XOR Data[46]) XOR (Data[28] OR Data[12]))) XOR ((Data[45] AND Data[4]) AND (NOT Data[31])))))))) XOR (((NOT (((NOT (NOT Data[19])) OR ((Data[30] OR (NOT ((Data[36] XOR Data[3]) XOR Data[50]))) AND Data[31])) AND Data[8])) XOR (((NOT (NOT (((Data[35] AND Data[23]) OR (Data[40] OR Data[11])) OR (((Data[12] XOR Data[42]) XOR Data[32]) OR (NOT Data[34]))))) AND (NOT Data[7])) AND ((Data[15] AND Data[27]) AND ((((NOT (((NOT Data[12]) XOR (NOT Data[21])) XOR (Data[39] OR Data[21]))) XOR ((NOT ((Data[31] XOR Data[26]) XOR Data[50])) OR ((((Data[7] XOR Data[6]) XOR Data[11]) XOR Data[18]) XOR Data[4]))) XOR ((((NOT Data[28]) AND ((Data[19] XOR Data[4]) XOR Data[16])) XOR (((NOT Data[23]) XOR ((Data[34] XOR Data[42]) XOR Data[15])) XOR ((Data[40] XOR Data[20]) XOR TRUE))) XOR ((NOT Data[6]) OR (Data[12] AND Data[2])))) OR (NOT ((Data[46] XOR ((Data[14] AND Data[43]) AND Data[50])) XOR Data[6])))))) XOR ((NOT (NOT (((Data[49] XOR ((Data[10] AND Data[41]) AND (FALSE AND Data[10]))) XOR ((((Data[38] XOR Data[33]) XOR Data[36]) XOR (Data[29] AND Data[4])) XOR Data[43])) AND (NOT ((NOT Data[3]) AND Data[9]))))) AND (NOT Data[5])))) XOR (((NOT ((NOT (((NOT Data[6]) AND (Data[1] OR Data[28])) AND (NOT ((Data[26] XOR Data[28]) XOR Data[16])))) AND (((NOT Data[18]) XOR Data[22]) XOR (((Data[20] AND Data[15]) OR (NOT Data[40])) AND (NOT (Data[2] AND Data[7])))))) OR (((((((Data[50] OR Data[5]) AND Data[50]) AND (((NOT Data[40]) XOR (Data[18] OR Data[38])) XOR (NOT Data[31]))) OR Data[48]) XOR (((((((Data[15] XOR Data[26]) XOR Data[23]) XOR (Data[33] OR Data[44])) XOR Data[6]) AND (NOT ((Data[35] XOR Data[26]) XOR Data[47]))) XOR (((NOT Data[7]) AND (NOT Data[14])) AND (Data[33] OR Data[50]))) XOR Data[48])) XOR (NOT (Data[32] OR (NOT (Data[20] OR Data[48]))))) AND (((((Data[16] OR (NOT Data[1])) OR (NOT (Data[46] AND Data[16]))) AND (((NOT Data[2]) OR (Data[36] AND Data[9])) OR ((Data[4] AND Data[34]) AND (Data[37] OR Data[13])))) XOR Data[23]) XOR (Data[4] OR (Data[27] OR (((Data[35] OR Data[31]) XOR (Data[9] OR Data[11])) XOR (Data[23] AND Data[37]))))))) AND (((Data[22] OR (((((NOT Data[32]) XOR ((Data[24] XOR Data[27]) XOR Data[47])) XOR Data[32]) OR ((NOT Data[37]) OR (NOT Data[46]))) AND Data[28])) AND (NOT (Data[8] OR (((NOT Data[42]) OR (Data[46] OR Data[24])) AND ((NOT Data[33]) AND ((Data[25] XOR Data[24]) XOR Data[9])))))) OR (((((Data[26] AND Data[8]) AND Data[49]) OR (NOT Data[2])) AND ((((Data[7] XOR ((Data[25] XOR Data[31]) XOR Data[21])) XOR (NOT Data[38])) OR ((Data[29] OR Data[14]) AND (Data[34] OR Data[25]))) AND ((NOT ((Data[18] XOR Data[6]) XOR Data[48])) AND Data[7]))) OR Data[13])))) XOR Data[37]) XOR (((NOT ((Data[15] XOR (NOT ((((NOT Data[46]) OR (Data[25] OR Data[41])) OR (((FALSE OR Data[14]) XOR ((Data[27] XOR Data[2]) XOR Data[33])) XOR (NOT Data[33]))) AND Data[17]))) XOR (Data[37] OR (((NOT ((Data[24] OR Data[45]) OR ((Data[33] XOR Data[46]) XOR Data[36]))) XOR (((NOT Data[10]) OR (Data[10] OR Data[28])) OR ((Data[3] OR Data[26]) AND Data[48]))) XOR (((Data[14] AND TRUE) AND (NOT Data[17])) OR ((NOT Data[50]) OR (Data[48] AND TRUE))))))) AND Data[17]) OR (((NOT ((((((Data[30] OR ((Data[12] OR Data[23]) AND Data[24])) XOR (((Data[13] XOR Data[11]) XOR Data[1]) OR (NOT Data[38]))) XOR (Data[39] AND (NOT ((Data[3] XOR Data[20]) XOR Data[5])))) XOR (Data[21] OR ((NOT (Data[33] OR Data[7])) OR Data[31]))) XOR (NOT (NOT Data[49]))) OR Data[41])) XOR ((TRUE XOR (((((Data[39] XOR ((((Data[17] AND Data[5]) AND Data[4]) XOR (NOT (Data[49] AND Data[25]))) XOR (NOT Data[39]))) XOR Data[32]) OR (NOT (Data[6] AND Data[44]))) XOR ((((Data[18] OR (NOT Data[31])) AND ((NOT Data[48]) OR (Data[21] OR Data[41]))) OR Data[20]) AND ((NOT ((NOT Data[28]) AND ((Data[18] XOR Data[44]) XOR Data[40]))) OR (Data[12] OR (((Data[5] OR Data[13]) XOR (Data[48] OR Data[34])) XOR Data[30]))))) XOR Data[23])) XOR Data[45])) XOR (((((NOT (NOT Data[44])) XOR ((((((FALSE XOR Data[24]) XOR Data[5]) OR ((Data[27] XOR Data[9]) XOR Data[19])) XOR ((Data[47] XOR ((Data[17] XOR Data[1]) XOR Data[11])) XOR Data[34])) XOR (NOT ((Data[23] XOR Data[47]) XOR Data[23]))) AND (((Data[7] OR ((Data[36] XOR TRUE) XOR Data[6])) XOR (((Data[5] XOR Data[2]) XOR Data[29]) OR ((Data[1] XOR Data[46]) XOR Data[47]))) XOR ((Data[40] AND Data[29]) AND ((Data[38] XOR Data[44]) XOR FALSE))))) XOR (((((Data[2] OR Data[12]) XOR (Data[1] OR Data[17])) XOR ((Data[17] XOR Data[4]) XOR Data[32])) OR (((Data[19] XOR Data[41]) XOR Data[36]) OR (Data[18] OR Data[5]))) OR Data[16])) OR (Data[45] OR (NOT ((Data[26] XOR (NOT (Data[22] AND Data[9]))) XOR ((Data[28] OR Data[40]) OR ((Data[39] XOR Data[15]) XOR Data[21])))))) AND (NOT (Data[24] OR ((((Data[38] OR Data[48]) OR (Data[8] AND Data[6])) AND ((((Data[38] XOR Data[9]) XOR Data[11]) XOR (Data[44] AND Data[3])) XOR (Data[11] OR Data[50]))) OR (((NOT Data[30]) AND (Data[37] AND Data[27])) OR ((NOT Data[5]) AND (Data[34] AND Data[22]))))))))));
    OutReady := 1;
    CollectInput(RESET:=TRUE);
  END_IF;
END_PROGRAM

CONFIGURATION Config0
  RESOURCE Res0 ON PLC
    TASK task0(INTERVAL := T#20ms,PRIORITY := 0);
    PROGRAM instance0 WITH task0 : Boiler;
  END_RESOURCE
END_CONFIGURATION
